(* IEC 61131-3 sources: daoli-st-library/DL_MathData (part 26) *)

(* ---- FC_DL_TimeDivChk.st ---- *)
(*
    FC_DL_TimeDivChk —— TIME 整数除法除零拦截与模长防御包装
    ------------------------------------------------------------------
    分类      : DL_MathData / TimeArith
    前缀      : FC_DL_
    版本      : 1.0.0
    溯源      : IEC 61131-3 标准语义的道莅防御性实现
                （内部委托平台内建函数，外围统一错误码/钳位/双语文档；
                  未复制任何闭源厂商源码，参考实现仅限 MIT/Apache 许可）
    平台      : 纯 IEC 61131-3，CODESYS / TwinCAT / InoProShop 通用
    作者      : 道莅代码库 · PLC编程专家（R16）
    ------------------------------------------------------------------
    功能说明  : TIME 整数除法：返回 tIn ÷ nDiv，TIME 算术委托 `÷` 运算符，
                不重实现任何时间运算内核；
                nDiv = 0 判为故障级 16#0001_02C7，返回 T#0S 且 bValid=FALSE（除零故障）；
                nDiv < 0 时取模长参与运算并置信息级 16#0001_01E6
                （TIME 无负语义，方向取模长，bError=FALSE、bValid=TRUE）；
                模长取负回绕防御：先将 INT 除子升位复制到 DINT 再取负，
                规避 INT 最小值 -32768 直接取负的回绕未定义行为；
                除法前已强制判定除子非零（nDiv = 0 分支提前拦截），满足除法前判除子红线；
                钳位方向：无钳位（除零故障拦截 / 负除子模长化记录）。
    错误码    : 16#0001_02C7 除数为 0（除零故障）——故障级，返回 T#0S
                16#0001_01E6 负除子输入，已按模长参与运算——信息级，正常防御
                16#0001_01E7 预留禁用（信息级，不得挪用）
                16#0001_02C8 预留禁用（故障级，不得挪用）
                16#0001_02C9 预留禁用（故障级，不得挪用）
    状态机    : R6 标注 N/A —— 本组件为纯函数无顺序状态机，无 CASE 可写，非法状态不可能出现，故以本节说明替代 ELSE 兜底
    修订记录  : 2026-11-16 v1.0.0 首次入库（R16）
*)
FUNCTION FC_DL_TimeDivChk : TIME
VAR_INPUT
    tIn  : TIME; // 输入时长（被除数） [ms] / input duration (dividend)
    nDiv : INT;  // 除子 [倍]，非 0，除零为故障 / divisor [x], nonzero, div-by-zero is a fault
END_VAR
VAR_OUTPUT
    eErr   : UDINT; // 错误码，0=正常 / error id, 0=ok
    bError : BOOL;  // 是否出错，eErr 非 0 时为 TRUE / error flag, TRUE when eErr is nonzero
    bValid : BOOL;  // 输出是否有效可用 / output valid flag
END_VAR
VAR CONSTANT
    DL_TIME_ZERO : TIME := T#0S; // TIME 零值（故障缺省返回） [ms] / TIME zero value (fault default return)
END_VAR
VAR
    nWiden : DINT; // 升位到 DINT 的除子副本 [倍] / divisor copy widened to DINT
    nAbs   : DINT; // 除子模长 [倍] / divisor magnitude
END_VAR

// 段 1｜返回值与错误状态预置 / segment 1, preset return value and error status
FC_DL_TimeDivChk := DL_TIME_ZERO; // 故障缺省返回 T#0S [ms] / fault default returns T#0S
eErr   := 0;     // 预置无错误 / preset no error
bError := FALSE; // 预置无故障 / preset no fault
bValid := FALSE; // 预置无效，通过除零闸后置位 / preset invalid, set TRUE after divide-by-zero guard

// 段 2｜除零故障闸 / segment 2, divide-by-zero fault guard
IF nDiv = 0 THEN
    FC_DL_TimeDivChk := DL_TIME_ZERO; // 故障级返回 T#0S [ms] / fault level returns T#0S
    eErr   := 16#0001_02C7;           // 除零故障码 / divide-by-zero fault id
    bError := TRUE;                   // 置故障标志 / set fault flag
    bValid := FALSE;                  // 输出无效 / output invalid
    RETURN;                           // 立即返回 / immediate return
END_IF

// 段 3｜除子模长整备（含取负回绕防御） / segment 3, divisor magnitude preparation with negation-wrap defense
nWiden := nDiv; // 先升位复制到 DINT / widen copy to DINT first
IF nDiv < 0 THEN
    nAbs := -nWiden; // DINT 域内取模长（规避 INT 最小值 -32768 取负回绕） / magnitude in DINT domain (avoids INT minimum -32768 negation wrap)
    eErr := 16#0001_01E6; // 信息级：负除子按模长处理（TIME 无负语义，方向取模长） / info level: negative divisor handled by magnitude (TIME has no negative semantics)
ELSE
    nAbs := nWiden; // 正除子模长即原值 / positive divisor, magnitude equals original
END_IF

// 段 4｜主体除法计算（末段） / segment 4, main division calculation (final)
FC_DL_TimeDivChk := tIn / nAbs; // 除子已判非零，模长参与委托 `÷` 运算符除法 / divisor checked nonzero, division via `÷` operator with magnitude
bError := FALSE; // 信息级模长化不置故障，除零分支已提前返回 / info-level magnitude never raises fault, divide-by-zero branch has returned
bValid := TRUE;  // 域内或模长化输出均有效可用 / in-domain or magnitude output is valid
END_FUNCTION

(* ---- FC_DL_TimeMulSat.st ---- *)
(*
    FC_DL_TimeMulSat —— TIME 整数乘法（乘数域闸 + 溢出饱和）
    ------------------------------------------------------------------
    分类      : DL_MathData / TimeArith
    前缀      : FC_DL_
    版本      : 1.0.0
    溯源      : IEC 61131-3 标准语义的道莅防御性实现
                （对照 IEC 61131-3 第 3 版 MUL_TIME 标准语义，委托平台内建 `*`
                  与 `/` 运算符，外围全部闸门 / 饱和 / 码位 / 双语文档 100% 自有；
                  clean-room 编写，未复制任何闭源厂商源码，参考实现仅限 MIT/Apache）
    平台      : 纯 IEC 61131-3，CODESYS 3.5 / TwinCAT 3 / InoProShop / Machine Expert 通用
    作者      : 道莅代码库 · PLC编程专家（R69 构建轮 · 批 1 · N1）
    ------------------------------------------------------------------
    功能说明  : TIME × 乘数。与库内既有 FC_DL_TimeScaleSat 的分工：ScaleSat 是
                「负乘子钳零、双乘子全放行」的宽松包装；本件是 MUL_TIME 的**严格域闸**
                版本——负乘子属于语义非法（时长无负语义）必须**禁入**并报故障级，
                乘数超 INT 正域上界（32767）同样禁入（防以超域乘子绕过溢出预判），
                只有域内合法乘子才进入乘法内核。
                溢出预判采用除法比较口径（R54 / 实战规则 6）：`tIn > MAX / nScale`，
                比较表达式中不出现乘 / 加运算符，命中即饱和夹 LTIME 上界并报信息级。
                乘数域上界反算依据（实战规则 9）：TIME 为 32 位毫秒容器
                （上限 4294967295 ms ≈ T#49D17H2M47S295MS），乘子上界取 32767（INT 正域）
                是为让 `MAX / nScale` 恒有整数解且不产生 0 除；乘子更大时预判式
                本身会因整数除法结果为 0 而把一切非零时长误判为溢出，故必须在域闸
                先行禁入，不得放大上界。
    错误码    : 16#0001_03F7 负乘子禁入（语义非法），输出 T#0S —— 故障级
                16#0001_03F8 乘子超上界 32767，输出 T#0S —— 故障级
                16#0001_04F6 乘法溢出，输出已饱和至 TIME 上界 —— 信息级，值可用
    码位总账  : 16#0001_03F7 / 03F8 用 ｜ 16#0001_04F6 用
    状态机    : R6 标注 N/A —— 纯函数无顺序状态机，无 CASE 可写，非法状态不可能出现
    采样约定  : 无定时器 / 无沿检测 / 无跨周期状态，结论与任务周期无关
    修订记录  : 2026-11-22 v1.0.0 首次入库（R69 构建轮 · 批 1 · N1）
*)
FUNCTION FC_DL_TimeMulSat : TIME
VAR_INPUT
    tIn     : TIME;                            // 被乘时长 [ms] / multiplicand duration [ms]
    diScale : DINT;                            // 乘数 [倍]，域 0..32767，负值与超上界禁入 / scale factor [x], domain 0..32767
END_VAR
VAR_OUTPUT
    eErr        : UDINT;                       // 错误码，0 = 正常 / error id, 0 = ok
    bError      : BOOL;                        // 故障标志，故障级码时为 TRUE / error flag, TRUE on fault level
    bValid      : BOOL;                        // 返回值可用（故障级为 FALSE）/ return usable, FALSE on fault level
    bSaturated  : BOOL;                        // 已饱和至 TIME 上界 / saturated at the TIME ceiling
END_VAR
VAR CONSTANT
    DL_TM_MAX   : TIME := T#49D17H2M47S295MS;  // 32 位 TIME 容器上限，等价 4294967295 ms [ms] / 32-bit TIME ceiling [ms]
    DL_TM_ZERO  : TIME := T#0S;                // TIME 零值（故障缺省返回） [ms] / TIME zero, the fault default
    DL_TM_SCALE_MAX : DINT := 32767;           // 乘数上界 [倍]，INT 正域上界（反算依据见头注释）/ scale ceiling [x]
    DL_TM_SCALE_MIN : DINT := 0;               // 乘数下界 [倍]，负值禁入 / scale floor [x]
END_VAR
VAR
    nScaleInt : INT;                           // 域内乘数（已过闸，可直接参与 TIME 运算）[倍] / in-domain scale as INT
END_VAR

// 段 1｜返回值与错误状态预置（实战规则 1① 四段式第一段）/ segment 1, preset return and status
FC_DL_TimeMulSat := DL_TM_ZERO;   // 故障缺省返回 T#0S [ms] / fault default returns T#0S
eErr       := 0;                  // 预置无错误 / preset no error
bError     := FALSE;              // 预置无故障 / preset no fault
bValid     := FALSE;              // 预置不可用，过闸后置位 / preset unusable, set TRUE after the gates
bSaturated := FALSE;              // 预置未饱和 / preset not saturated

// 段 2｜乘数域闸：负值禁入（语义非法）/ segment 2, scale domain gate, negative is refused
IF diScale < DL_TM_SCALE_MIN THEN
    eErr   := 16#0001_03F7;       // 故障级：负乘子禁入 / fault level: negative factor refused
    bError := TRUE;               // R45 配对置故障标志 / raise the error flag, paired with the code
    bValid := FALSE;              // 返回值不可用 / return unusable
    RETURN;                       // 出口，不触碰乘法内核 / exit, the kernel is never touched
END_IF

// 段 3｜乘数域闸：超上界禁入（防以超域乘子绕过溢出预判）/ segment 3, upper domain gate
IF diScale > DL_TM_SCALE_MAX THEN
    eErr   := 16#0001_03F8;       // 故障级：乘子超上界 / fault level: factor above the ceiling
    bError := TRUE;               // R45 配对 / paired with the code
    bValid := FALSE;              // 返回值不可用 / return unusable
    RETURN;                       // 出口 / exit
END_IF
nScaleInt := DINT_TO_INT(diScale);   // 域内乘数降为 INT（域已证 <= 32767，无窄化风险）[倍] / in-domain scale to INT

// 段 4｜零乘子：合法零乘，输出 T#0S 且无码（零乘不是错误）/ segment 4, legal zero multiply
IF nScaleInt = 0 THEN
    FC_DL_TimeMulSat := DL_TM_ZERO;   // 零乘结果 [ms] / zero product
    bValid := TRUE;                   // 零是可用结果 / zero is a usable result
    RETURN;                           // 出口 / exit
END_IF

// 段 5｜溢出预判（除法比较口径）+ 域内委托乘法内核 / segment 5, divide-compare pre-check then delegate
IF tIn > (DL_TM_MAX / nScaleInt) THEN
    FC_DL_TimeMulSat := DL_TM_MAX;    // 预判命中：饱和夹上界（除子 nScaleInt > 0 恒非零）[ms] / saturate to the ceiling
    eErr       := 16#0001_04F6;       // 信息级：乘法溢出已饱和 / info level: overflow saturated
    bSaturated := TRUE;               // 饱和标志供上层计量 / saturation flag for the caller
ELSE
    FC_DL_TimeMulSat := tIn * nScaleInt;   // 域内委托 `*` 运算符内核 [ms] / in-domain multiplication kernel
END_IF
bError := FALSE;   // 信息级饱和不置故障（饱和是防御而非故障）/ info-level saturation is a defence, not a fault
bValid := TRUE;    // 域内或饱和输出均可用 / usable in the in-domain and the saturated path
END_FUNCTION

(* ---- FC_DL_TimeRatioCalc.st ---- *)
(*
    FC_DL_TimeRatioCalc —— 两个 TIME 的无量纲比值
    ------------------------------------------------------------------
    分类      : DL_MathData / Convert
    前缀      : FC_DL_
    版本      : 1.0.0
    溯源      : 公开算术定义的道莅防御性实现（比值 = 分子时长 / 分母时长）；
                库内 FC_DL_TimeDivChk 只出整数毫秒商（小数全丢），本件用 LREAL 承载
                以保留 15 位有效数字；饱和限、取模长口径、错误分级、双语文档 100% 自有；
                clean-room 重写，未复制任何闭源厂商源码，参考实现仅限 MIT/Apache 许可
    平台      : 纯 IEC 61131-3，CODESYS V3.5+ / TwinCAT 3 / InoProShop 通用
    作者      : 道莅代码库 · PLC编程专家（R19）
    ------------------------------------------------------------------
    功能说明  : 计算节拍分析 / 稼动率 / 循环时间偏差 / 加速比所需的比值，可选 ×100 出百分比。
                核心防御：① 分母毫秒值为 0 是除零唯一出口（故障级 0321 早退，绝不进入除法）；
                ② 分母模长 < 1 ms 视为无意义分母，比值直接饱和到 fRatioSpan（1 ms 以下
                   的分母在任何现场都无意义，且会让比值爆炸）；
                ③ 输入为负时按模长参与运算（TIME 的平台符号语义不一致，方向差异
                   由本件统一吃掉），并置信息码 0402；
                ④ 比值超 fRatioSpan 双侧钳位，禁 NaN / ±INF 穿透；
                ⑤ 同一拍同时命中两条信息级时以 0403（饱和）为准，码位单值不可并列。
                职责边界：本件只出比值，不做时间加减、不做时基换算。
    错误码    : 16#0001_0402 分母模长 < 1 ms 或输入为负，已按模长运算/饱和——信息级，正常防御
                16#0001_0403 比值超 fRatioSpan 已钳位（bSaturated = TRUE）——信息级，正常防御
                16#0001_0321 分母为 0（除零）——故障级，返回 0.0 且 bValid = FALSE
                16#0001_0322 结果非有限（NaN / ±INF）或比值上限参数非法——故障级，返回 0.0
                16#0001_0323 预留禁用（故障级，不得挪用）
    码位总账  : 16#0001_0402 用 / 16#0001_0403 用 ｜ 16#0001_0321 用 / 16#0001_0322 用 / 16#0001_0323 预留
    状态机    : R6 标注 N/A —— 本组件为纯函数无顺序状态机，无 CASE 可写，非法状态不可能出现
    采样约定  : 本件无定时器、无沿检测；TIME 实参由调用方按自身时基给出，结论与任务周期无关。
    修订记录  : 2026-11-16 v1.0.0 首次入库（R19）
*)
FUNCTION FC_DL_TimeRatioCalc : LREAL
VAR_INPUT
    tNumerator      : TIME := T#0S;           // 分子时长 [ms]，域 -24 h~+24 h / numerator duration [ms], domain -24 h~+24 h
    tDenominator    : TIME := T#1S;           // 分母时长 [ms]，域 -24 h~+24 h，模长须 ≥ 1 ms / denominator duration [ms], domain -24 h~+24 h, magnitude >= 1 ms
    bAsPercent      : BOOL := FALSE;          // TRUE = 结果 ×100 输出百分比 [%] / TRUE multiplies the result by 100 to percent [%]
    fRatioSpan      : LREAL := 1.0E6;         // 比值饱和上限（作用在返回量上）[无量纲]，域 1.0~1.0E12 / ratio saturation span applied to the returned value [dimensionless], 1.0~1.0E12
END_VAR
VAR_OUTPUT
    eErr            : UDINT;                  // 错误码，0=正常 / error id, 0=ok
    bError          : BOOL;                   // 故障标志，eErr 为故障级时 TRUE / error flag, TRUE on fault-level eErr
    bValid          : BOOL;                   // 返回值是否可用 / return value valid flag
    fRatioAbs       : LREAL;                  // 比值绝对值（HMI 只看量级用）[无量纲] / absolute ratio for HMI magnitude view [dimensionless]
    bSaturated      : BOOL;                   // 比值已饱和到 fRatioSpan / ratio saturated to fRatioSpan
END_VAR
VAR CONSTANT
    DL_FLOAT_EPS        : REAL := 1.0E-6;     // 浮点判等容差 [无量纲] / float equality tolerance [dimensionless]
    DL_TR_MIN_DEN_MS    : LREAL := 1.0;       // 分母模长下限 [ms] / denominator magnitude lower bound [ms]
    DL_TR_PERCENT       : LREAL := 100.0;     // 百分比放大因子 [无量纲] / percent scale factor [dimensionless]
    DL_TR_SPAN_MIN      : LREAL := 1.0;       // 比值上限最小值 [无量纲] / minimum ratio span [dimensionless]
    DL_TR_SPAN_MAX      : LREAL := 1.0E12;    // 比值上限最大值 [无量纲] / maximum ratio span [dimensionless]
    DL_TR_INF_GUARD     : LREAL := 1.0E300;   // 非有限幅值判定阈值 [无量纲] / non-finite magnitude guard [dimensionless]
    DL_TR_ZERO          : LREAL := 0.0;       // 零值常量，避免裸字面量 [无量纲] / zero constant, avoids a bare literal [dimensionless]
END_VAR
VAR
    fNumAbs         : LREAL;                  // 分子模长 [ms] / numerator magnitude [ms]
    fDenAbs         : LREAL;                  // 分母模长 [ms] / denominator magnitude [ms]
    fSpanEff        : LREAL;                  // 生效比值上限，钳位后使用 [无量纲] / effective ratio span after clamping [dimensionless]
    fRatio          : LREAL;                  // 计算中的比值中间量 [无量纲] / ratio intermediate value [dimensionless]
    nDenMs          : DINT;                   // 分母毫秒整数形态，除零判定用 [ms] / denominator in integer milliseconds, used for the divide-by-zero gate [ms]
    bNegativeIn     : BOOL;                   // 输入存在负值时基的标志 / flag for negative time base inputs
END_VAR

// 段 1｜返回值与错误状态预置 / segment 1, preset return value and error status
FC_DL_TimeRatioCalc := DL_TR_ZERO;            // 故障缺省返回 0.0 / fault default returns zero
eErr := 0;                                    // 预置无错误 / preset no error
bError := FALSE;                              // 预置无故障 / preset no fault
bValid := FALSE;                              // 预置不可用，通过闸门后置位 / preset invalid, set TRUE after the gates
fRatioAbs := DL_TR_ZERO;                      // 量级输出先清零 / clear the magnitude output
bSaturated := FALSE;                          // 预置未饱和 / preset not saturated

// 段 2｜比值上限参数闸（非法上限等于比值域不存在，落入结果不可表示）/ segment 2, ratio span gate
fSpanEff := fRatioSpan;                       // 取入参副本，不改调用方数据 / copy the input, never modify caller data
IF (fSpanEff <> fSpanEff) OR (fSpanEff > DL_TR_INF_GUARD) OR (fSpanEff < -DL_TR_INF_GUARD) THEN
    eErr := 16#0001_0322;                     // 上限非有限即结果不可表示 / a non-finite span makes the result unrepresentable
    bError := TRUE;                           // 置故障标志 / raise the error flag
    RETURN;                                   // 故障级提前返回 / early return on fault
END_IF
IF fSpanEff < DL_TR_SPAN_MIN THEN
    fSpanEff := DL_TR_SPAN_MIN;               // 上限过小钳到 1.0，避免比值域退化 / clamp a too small span to 1.0
    eErr := 16#0001_0403;                     // 信息级：上限已钳位 / info level, the span has been clamped
ELSIF fSpanEff > DL_TR_SPAN_MAX THEN
    fSpanEff := DL_TR_SPAN_MAX;               // 上限过大钳到 1.0E12 / clamp an oversized span to 1.0E12
    eErr := 16#0001_0403;                     // 信息级：上限已钳位 / info level, the span has been clamped
END_IF

// 段 3｜除零唯一出口（先取整数毫秒判定，再进入浮点除法）/ segment 3, the only divide-by-zero exit
nDenMs := TIME_TO_DINT(tDenominator);         // 显式取分母毫秒整数，禁隐式换算 / take denominator milliseconds explicitly, no implicit cast
IF nDenMs = 0 THEN
    eErr := 16#0001_0321;                     // 除零故障码 / divide-by-zero fault id
    bError := TRUE;                           // 置故障标志 / raise the error flag
    bValid := FALSE;                          // 结果不可用 / result not usable
    RETURN;                                   // 故障级提前返回，绝不进入除法 / early return, the division is never executed
END_IF

// 段 4｜按模长参与运算（TIME 符号语义跨平台不一致，方向差异在此统一吃掉）/ segment 4, magnitudes only
fNumAbs := ABS(TIME_TO_LREAL(tNumerator));    // 分子模长 [ms] / numerator magnitude [ms]
fDenAbs := ABS(TIME_TO_LREAL(tDenominator));  // 分母模长 [ms] / denominator magnitude [ms]
bNegativeIn := (TIME_TO_DINT(tNumerator) < 0) OR (nDenMs < 0); // 负时基判定 / negative time base detection
IF bNegativeIn THEN
    eErr := 16#0001_0402;                     // 信息级：输入为负已按模长运算 / info level, negative inputs are handled by magnitude
END_IF

// 段 5｜分母过小闸：不足 1 ms 直接饱和，不做除法 / segment 5, tiny-denominator gate
IF fDenAbs < DL_TR_MIN_DEN_MS THEN
    fRatio := fSpanEff;                       // 过小分母直接给饱和值，规避比值爆炸 / jump straight to the span, avoid an exploding ratio
    bSaturated := TRUE;                       // 标记饱和 / flag the saturation
    eErr := 16#0001_0402;                     // 信息级：分母过小已饱和 / info level, tiny denominator saturated
ELSE
    fRatio := fNumAbs / fDenAbs;              // 分母模长 ≥ 1 ms，除法安全 / the denominator is at least 1 ms, the division is safe
    IF bAsPercent THEN
        fRatio := fRatio * DL_TR_PERCENT;     // 可选百分比放大 [%] / optional percent scaling [%]
    END_IF
END_IF

// 段 6｜结果非有限复检（NaN 穿透拦截）/ segment 6, non-finite recheck
IF (fRatio <> fRatio) OR (fRatio > DL_TR_INF_GUARD) OR (fRatio < -DL_TR_INF_GUARD) THEN
    eErr := 16#0001_0322;                     // 结果非有限故障码 / non-finite result fault id
    bError := TRUE;                           // 置故障标志 / raise the error flag
    bValid := FALSE;                          // 结果不可用 / result not usable
    FC_DL_TimeRatioCalc := DL_TR_ZERO;        // 明确返回 0.0 / return zero explicitly
    RETURN;                                   // 故障级提前返回 / early return on fault
END_IF

// 段 7｜饱和钳位（单侧上限，比值恒非负）/ segment 7, saturation clamp
IF fRatio > fSpanEff THEN
    fRatio := fSpanEff;                       // 钳到生效上限 / clamp to the effective span
    bSaturated := TRUE;                       // 标记饱和 / flag the saturation
    eErr := 16#0001_0403;                     // 信息级：超上限已钳位，与 0402 同拍时以本码为准 / info level, clamped; this id wins over 0402 in the same cycle
END_IF

// 段 8｜发布结果 / segment 8, publish the result
FC_DL_TimeRatioCalc := fRatio;                // 输出比值（含百分比放大） [无量纲] / publish the ratio incl. percent scaling [dimensionless]
fRatioAbs := fRatio;                          // 比值恒按模长运算，量级即本身 / the ratio is magnitude based, so the magnitude equals the value
bValid := TRUE;                               // 通过全部闸门，结果可用 / all gates passed, the result is usable
bError := FALSE;                              // 信息级不置故障 / info level never raises a fault
END_FUNCTION

(* ---- FC_DL_TimeScaleSat.st ---- *)
(*
    FC_DL_TimeScaleSat —— TIME 整数乘法溢出饱和防御包装
    ------------------------------------------------------------------
    分类      : DL_MathData / TimeArith
    前缀      : FC_DL_
    版本      : 1.0.0
    溯源      : IEC 61131-3 标准语义的道莅防御性实现
                （内部委托平台内建函数，外围统一错误码/钳位/双语文档；
                  未复制任何闭源厂商源码，参考实现仅限 MIT/Apache 许可）
    平台      : 纯 IEC 61131-3，CODESYS / TwinCAT / InoProShop 通用
    作者      : 道莅代码库 · PLC编程专家（R16）
    ------------------------------------------------------------------
    功能说明  : TIME 整数乘法：返回 tIn × nScale，TIME 算术委托 `×` 运算符，
                不重实现任何时间运算内核；
                nScale < 0 时防御性输出 T#0S 并置信息级 16#0001_01E5
                （TIME 无负语义，负乘子按钳零处理，bError=FALSE、bValid=TRUE）；
                nScale = 0 时输出 T#0S，无错误码（零乘合法）；
                溢出预判采用除法比较口径（规避「先算后判」红线）：
                nScale > 0 且 tIn > DL_TIME_MAX / nScale 时判乘法将溢出，
                直接饱和输出 DL_TIME_MAX，置信息级 16#0001_01E4；
                预判除法除子 nScale > 0 恒非零，满足除法前判除子红线；
                钳位方向：负乘子钳零 / 正乘子溢出钳上界 DL_TIME_MAX（双侧饱和语义）。
    错误码    : 16#0001_01E4 乘法结果超 TIME 上限，已饱和至 DL_TIME_MAX——信息级，正常防御
                16#0001_01E5 负乘子输入，已钳位输出 T#0S——信息级，正常防御
                16#0001_02C4 预留禁用（故障级，不得挪用）
                16#0001_02C5 预留禁用（故障级，不得挪用）
                16#0001_02C6 预留禁用（故障级，不得挪用）
    状态机    : R6 标注 N/A —— 本组件为纯函数无顺序状态机，无 CASE 可写，非法状态不可能出现，故以本节说明替代 ELSE 兜底
    修订记录  : 2026-11-16 v1.0.0 首次入库（R16）
*)
FUNCTION FC_DL_TimeScaleSat : TIME
VAR_INPUT
    tIn    : TIME; // 输入时长 [ms] / input duration
    nScale : INT;  // 乘子 [倍]，0~32767，负值输出钳 T#0s / scale factor [x], 0~32767, negative clamps output to T#0s
END_VAR
VAR_OUTPUT
    eErr   : UDINT; // 错误码，0=正常 / error id, 0=ok
    bError : BOOL;  // 是否出错，eErr 非 0 时为 TRUE / error flag, TRUE when eErr is nonzero
    bValid : BOOL;  // 输出是否有效可用 / output valid flag
END_VAR
VAR CONSTANT
    DL_TIME_MAX  : TIME := T#49D17H2M47S295MS; // 32 位 TIME 容器上限，等价 4294967295 ms [ms] / 32-bit TIME container ceiling, equals 4294967295 ms
    DL_TIME_ZERO : TIME := T#0S;               // TIME 零值（钳位目标） [ms] / TIME zero value (clamp target)
END_VAR

// 段 1｜返回值与错误状态预置 / segment 1, preset return value and error status
FC_DL_TimeScaleSat := DL_TIME_ZERO; // 故障缺省返回 T#0S [ms] / fault default returns T#0S
eErr   := 0;     // 预置无错误 / preset no error
bError := FALSE; // 预置无故障（本组件无故障级路径） / preset no fault (no fault-level path in this component)
bValid := FALSE; // 预置无效，通过乘子判定后置位 / preset invalid, set TRUE after factor check

// 段 2｜乘子符号判定 / segment 2, scale factor sign check
IF nScale < 0 THEN
    FC_DL_TimeScaleSat := DL_TIME_ZERO; // 负乘子钳位输出 T#0S（TIME 无负语义） / negative factor clamps output to T#0S (TIME has no negative semantics)
    eErr := 16#0001_01E5;               // 信息级：负乘子已钳零 / info level: negative factor clamped to zero
    bError := FALSE;                    // 信息级钳零不置故障 / info-level clamp never raises fault
    bValid := TRUE;                     // 钳零输出有效可用 / clamped output is valid
    RETURN;                             // 立即返回 / immediate return
ELSIF nScale = 0 THEN
    FC_DL_TimeScaleSat := DL_TIME_ZERO; // 零乘子输出 T#0S（零乘合法，无错误码） / zero factor yields T#0S (legal zero multiply, no error id)
    bError := FALSE;                    // 无故障 / no fault
    bValid := TRUE;                     // 输出有效可用 / output is valid
    RETURN;                             // 立即返回 / immediate return
END_IF

// 段 3｜除法比较溢出预判与主体乘法（末段） / segment 3, divide-compare overflow pre-check and main multiplication (final)
IF tIn > DL_TIME_MAX / nScale THEN
    FC_DL_TimeScaleSat := DL_TIME_MAX; // 溢出预判命中，饱和至上限（除子 nScale > 0 恒非零） / overflow pre-check hit, saturate to ceiling (divisor nScale > 0 guaranteed nonzero)
    eErr := 16#0001_01E4;              // 信息级：乘法溢出已饱和 / info level: multiplication overflow, saturated
ELSE
    FC_DL_TimeScaleSat := tIn * nScale; // 预判通过，域内委托 `×` 运算符乘法 / pre-check passed, in-domain multiplication via `×` operator
    eErr := 0; // 域内无错误 / in-domain, no error
END_IF
bError := FALSE; // 信息级饱和不置故障 / info-level saturation never raises fault
bValid := TRUE;  // 域内或饱和输出均有效可用 / in-domain or saturated output is valid
END_FUNCTION

(* ---- FC_DL_TimeSubSat.st ---- *)
(*
    FC_DL_TimeSubSat —— TIME 减法负差钳零防御包装
    ------------------------------------------------------------------
    分类      : DL_MathData / TimeArith
    前缀      : FC_DL_
    版本      : 1.0.0
    溯源      : IEC 61131-3 标准语义的道莅防御性实现
                （内部委托平台内建函数，外围统一错误码/钳位/双语文档；
                  未复制任何闭源厂商源码，参考实现仅限 MIT/Apache 许可）
    平台      : 纯 IEC 61131-3，CODESYS / TwinCAT / InoProShop 通用
    作者      : 道莅代码库 · PLC编程专家（R16）
    ------------------------------------------------------------------
    功能说明  : TIME 减法：返回 tA - tB（tA 为被减数、tB 为减数），TIME 算术
                委托 `-` 运算符，不重实现任何时间运算内核；
                tB > tA 时差为负，而 TIME 为无符号语义、负差跨平台未定义，
                故防御性钳位输出 T#0S 并置信息级 16#0001_01E2
                （bError=FALSE、bValid=TRUE，属正常防御）；
                钳位方向：仅下界单侧钳零（负差归 T#0S，不产生回绕）；
                本组件无故障级路径（减法运算不存在除法/非有限态故障源），
                故障三码位预留禁用。
    错误码    : 16#0001_01E2 减数为大，负差已钳位至 T#0S——信息级，正常防御
                16#0001_01E3 预留禁用（信息级，不得挪用）
                16#0001_02C1 预留禁用（故障级，不得挪用）
                16#0001_02C2 预留禁用（故障级，不得挪用）
                16#0001_02C3 预留禁用（故障级，不得挪用）
    状态机    : R6 标注 N/A —— 本组件为纯函数无顺序状态机，无 CASE 可写，非法状态不可能出现，故以本节说明替代 ELSE 兜底
    修订记录  : 2026-11-16 v1.0.0 首次入库（R16）
*)
FUNCTION FC_DL_TimeSubSat : TIME
VAR_INPUT
    tA : TIME; // 被减数 [ms] / minuend
    tB : TIME; // 减数 [ms] / subtrahend
END_VAR
VAR_OUTPUT
    eErr   : UDINT; // 错误码，0=正常 / error id, 0=ok
    bError : BOOL;  // 是否出错，eErr 非 0 时为 TRUE / error flag, TRUE when eErr is nonzero
    bValid : BOOL;  // 输出是否有效可用 / output valid flag
END_VAR
VAR CONSTANT
    DL_TIME_ZERO : TIME := T#0S; // TIME 零值（负差钳位目标） [ms] / TIME zero value (clamp target for negative difference)
END_VAR

// 段 1｜返回值与错误状态预置 / segment 1, preset return value and error status
FC_DL_TimeSubSat := DL_TIME_ZERO; // 故障缺省返回 T#0S [ms] / fault default returns T#0S
eErr   := 0;     // 预置无错误 / preset no error
bError := FALSE; // 预置无故障（本组件无故障级路径） / preset no fault (no fault-level path in this component)
bValid := FALSE; // 预置无效，通过负差判定后置位 / preset invalid, set TRUE after negative-difference check

// 段 2｜负差钳零判定与主体减法（末段） / segment 2, negative-difference clamp-to-zero check and main subtraction (final)
IF tB > tA THEN
    FC_DL_TimeSubSat := DL_TIME_ZERO; // 负差钳位至 T#0S（TIME 无符号语义，负差跨平台未定义） / negative difference clamped to T#0S (TIME is unsigned, negative difference is platform-undefined)
    eErr := 16#0001_01E2;             // 信息级：负差已钳零 / info level: negative difference clamped to zero
ELSE
    FC_DL_TimeSubSat := tA - tB; // 域内委托 `-` 运算符减法 / in-domain subtraction via `-` operator
    eErr := 0; // 域内无错误 / in-domain, no error
END_IF
bError := FALSE; // 信息级钳零不置故障 / info-level clamp never raises fault
bValid := TRUE;  // 域内或钳零输出均有效可用 / in-domain or clamped output is valid
END_FUNCTION

(* ---- FC_DL_TimeToDintMs.st ---- *)
(*
    FC_DL_TimeToDintMs —— TIME 到 DINT 毫秒防御转换（超域饱和）
    ------------------------------------------------------------------
    分类      : DL_MathData / TimeConv
    前缀      : FC_DL_
    版本      : 1.0.0
    溯源      : IEC 61131-3 标准语义的道莅防御性实现
                （接口语义由 IEC 61131-3 定义，内部委托平台内建 TIME_TO_DINT，
                  外围统一错误码 / 钳位 / 双语文档；clean-room 重写，
                  未复制任何闭源厂商源码，参考实现仅限 MIT/Apache 许可）
    平台      : 纯 IEC 61131-3，CODESYS / TwinCAT / InoProShop 通用
    作者      : 道莅代码库 · PLC编程专家（R17）
    ------------------------------------------------------------------
    功能说明  : 将 TIME 值防御性转换为 DINT 毫秒数并作为返回值输出，域内委托平台内建 TIME_TO_DINT；
                溢出预判先行：先在 TIME 域与 2147483647 ms（T#24D20H31M23S647MS）比较，
                超限直接饱和输出 2147483647 并置信息级 16#0001_01F2，
                严禁把超限值送进 TIME_TO_DINT（部分平台此时返回负值，静默翻转语义）；
                转换结果为负（负 TIME 或平台回绕）时钳 0 并置信息级 16#0001_01F3；
                钳位方向：上界饱和至 2147483647 ms，下界钳 0 ms；
                纯值类型域无 NaN/±INF 态，故无故障级路径（三个故障槽预留）。
    错误码    : 16#0001_01F2 输入超 DINT 毫秒域（> 2147483647 ms），已饱和——信息级，正常防御
                16#0001_01F3 转换结果为负（负 TIME 或平台回绕），已钳 0——信息级，正常防御
                16#0001_02D9 预留禁用（故障级，不得挪用）
                16#0001_02DA 预留禁用（故障级，不得挪用）
                16#0001_02DB 预留禁用（故障级，不得挪用）
    状态机    : R6 标注 N/A —— 本组件为纯函数无顺序状态机，无 CASE 可写，非法状态不可能出现，故以本节说明替代 ELSE 兜底
    修订记录  : 2026-11-16 v1.0.0 首次入库（R17）
*)
FUNCTION FC_DL_TimeToDintMs : DINT
VAR_INPUT
    tIn : TIME; // 待转换时间值，有效域 0 ms ~ 4294967295 ms [ms] / time value to convert, domain 0 ms .. 4294967295 ms [ms]
END_VAR
VAR_OUTPUT
    eErr   : UDINT; // 错误码，0=正常 / error id, 0=ok
    bError : BOOL;  // 是否出错，eErr 非 0 时为 TRUE / error flag, TRUE when eErr is nonzero
    bValid : BOOL;  // 输出是否有效可用 / output valid flag
END_VAR
VAR CONSTANT
    DL_TIME_DINT_MAX : TIME := T#24D20H31M23S647MS; // DINT 正域可承载的最大毫秒数 2147483647 ms [ms] / max ms a DINT can carry, 2147483647 ms [ms]
    DL_DINT_MAX_MS   : DINT := 2147483647;          // 上界饱和输出值 [ms] / upper saturation output [ms]
    DL_MS_MIN        : DINT := 0;                   // 下界钳位值（TIME 无负语义） [ms] / lower clamp, TIME has no negative semantics [ms]
END_VAR
VAR
    nOut : DINT; // 域内转换中间结果 [ms] / in-domain conversion intermediate [ms]
END_VAR

// 段 1｜返回值与错误状态预置 / segment 1, preset return value and error status
FC_DL_TimeToDintMs := DL_MS_MIN; // 故障缺省返回 0 ms（TIME 无负语义） [ms] / fault default 0 ms, TIME has no negative semantics [ms]
eErr   := 0;     // 预置无错误 / preset no error
bError := FALSE; // 预置无故障（本件无故障级路径） / preset no fault, no fault-level path here
bValid := FALSE; // 预置输出无效，通过上界预判后置位 / preset invalid, set TRUE after the upper-bound pre-check

// 段 2｜上界预判与饱和（先判后算，禁先转换） / segment 2, upper bound pre-check and saturation (compare before convert)
IF tIn > DL_TIME_DINT_MAX THEN // 在 TIME 域先比较，绝不让超限值进入内建转换 [ms] / compare in the TIME domain first, never let an oversized value reach the built-in conversion [ms]
    FC_DL_TimeToDintMs := DL_DINT_MAX_MS; // 饱和输出 DINT 正域上限 2147483647 ms [ms] / saturate to the DINT positive bound 2147483647 ms [ms]
    eErr := 16#0001_01F2;                 // 信息级：超 DINT 毫秒域已饱和，正常防御 / info level: beyond the DINT ms domain, saturated
    bError := FALSE;                      // 信息级不置故障 / info level never raises fault
    bValid := TRUE;                       // 饱和值本身有效可用 / the saturated value itself is valid
    RETURN;                               // 饱和即出口，不调用内建转换 / saturation is the exit, built-in conversion not called
END_IF

// 段 3｜域内委托转换与负值钳零（末段） / segment 3, in-domain delegated conversion and negative clamp (final)
nOut := TIME_TO_DINT(tIn); // 域内委托平台内建 TIME_TO_DINT [ms] / in-domain delegate to built-in TIME_TO_DINT [ms]
IF nOut < DL_MS_MIN THEN
    nOut := DL_MS_MIN;    // 负结果钳 0（负 TIME 或平台回绕，TIME 无负语义） [ms] / clamp negative results to 0, TIME has no negative semantics [ms]
    eErr := 16#0001_01F3; // 信息级：结果为负已钳零，正常防御 / info level: result was negative and clamped to zero
ELSE
    eErr := 0;            // 域内无错误 / in-domain, no error
END_IF
FC_DL_TimeToDintMs := nOut; // 输出钳位后的毫秒结果 [ms] / output the clamped millisecond result [ms]
bError := FALSE;            // 信息级不置故障 / info level never raises fault
bValid := TRUE;             // 域内或钳位后输出均有效可用 / in-domain or clamped output is valid
END_FUNCTION

(* ---- FC_DL_TimeToHmsString.st ---- *)
(*
    组件名称 : FC_DL_TimeToHmsString
    所属子库 : DL_MathData
    当前版本 : 1.0.0
    兼 容 性 : CODESYS V3.5+ / TwinCAT 3 / 汇川 InoProShop；仅依赖 Standard.library
    功能描述 : TIME 时长 → 'HH:MM:SS.mmm' 定宽文本，负时长统一带负号，并把总小时数单独出口供报表使用。
              取舍 ①：不委托 DINT_TO_STRING 补零 —— 各平台对「正数是否带前导空格」「负数符号位置」
              的实现互不相同（R79 家族），靠它拼定宽字段必出「_1:05:03」这类带空格的串。
              本件用数字字符表 MID 取值 + CONCAT 拼装，位数与字符完全由代码控制。
              取舍 ②：负数先取绝对值再分解，但 DINT_MIN 单独走哨兵分支 —— −(−2147483648) 在 DINT 域回绕成自身，
              直接取负会把「最大负时长」变成「最大正时长」且符号丢失；本件对下界显式夹到 DINT_MAX 并保留负号。
              取舍 ③：分解全程只用非负操作数 —— 取绝对值之后再 MOD/DIV，三平台的负数取余歧义从源头消失。
              取舍 ④：小时字段不设上限截断，只发宽度提示 —— TIME 上限约 596 小时，HMI 常见 2 位小时字段装不下，
              但截断小时会让时长错得无声无息，宁可超宽 + 信息码让上位机改字段宽度。
    开源溯源 : T2-1 LGF Converter 子族（只借「时长转定宽文本」这一行为定义）。码位、补零策略、负数口径、；本件为道莅 clean-room 防御性实现（仅借 LGF 分类事实/参数域/行为定义，零代码行与符号名复制）。
              分解顺序 100% 自有，零代码行与注释复制。
    本文件内含 : FUNCTION FC_DL_TimeToHmsString（单 POU，无配套类型）
    依 赖 : 无 DL_ 内部依赖；Standard.library: LEN / MID / CONCAT
    红线自检 : R1 ✓ 零全局变量与外部变量 ｜ R2 ✓ 零物理 IO 地址
              R3 ✓ 纯 IEC 61131-3 ｜ R4 ✓ 下界哨兵 + 小时域闸 + 分解操作数恒非负 + 输出长度自证
              R5 ✓ 全变量中英双语同行注释 ｜ R6 N/A 纯函数无顺序状态机，无 CASE 可写
              R7 N/A 无定时器、无沿检测实例 ｜ R8 ✓ 毫秒基数、字段宽度、小时上限全常量化
    错误码   : 16#0001_044E [信息级] 负时长已带负号输出，bValid = TRUE
               16#0001_044F [信息级] 小时超 99，HMI 两位小时字段装不下，bValid = TRUE
               16#0001_0393 [故障级] 分解中间量非法（小时超 999，理论不可达），返回 '00:00:00.000'，bValid = FALSE
               16#0001_0394 [故障级] 预留禁用（不得挪用）
               16#0001_0395 [故障级] 预留禁用（不得挪用）
    码位总账 : 16#0001_044E 用 / 16#0001_044F 用 ｜ 16#0001_0393 用 / 16#0001_0394 预留 / 16#0001_0395 预留
    遗留假设 : ① 本件依赖「平台 TIME 为 32 位有符号毫秒计数」这一口径（TIME_TO_DINT 与 TIME 同宽）。
              CODESYS / TwinCAT 3 默认如此，InoProShop 未实测；若某平台 TIME 换成 64 位 LTime 语义，
              小时上限与 DINT_MIN 哨兵都需重估。交付门槛：三平台各编译并跑 T#-1ms、T#-2147483648ms、
              T#596H 三个边界 —— 未实测，编译门槛未闭合。
              ② MID 参数序按 IEC 标准 MID(串, 长度, 位置)，与库内既有用法同序。
    修订历史 :
        2026-11-16  v1.0.0  首版，R21 批次 3 入库
*)
FUNCTION FC_DL_TimeToHmsString : STRING
VAR_INPUT
    tIn             : TIME;   // 待格式化时长，全域（含负值）[ms] / duration to format, negative values included [ms]
END_VAR
VAR_OUTPUT
    eErr            : UDINT;  // 错误码，0=正常；16#0001_04XX 信息级 / 16#0001_03XX 故障级 / error id, 0=ok
    bError          : BOOL;   // 故障级标志，eErr 落 16#0001_03XX 时为 TRUE / fault flag, TRUE on fault-level eErr
    bValid          : BOOL;   // 返回值是否可用 / result usable flag
    bNegative       : BOOL;   // 输入是否为负时长，输出串因此带前导负号 / TRUE when the input duration is negative and the text carries a minus sign
    nTotalHours     : DINT;   // 总小时数（分解后），供报表直接取用 [h] / total hours after the decomposition [h]
END_VAR
VAR
    nMs             : DINT;   // 时长的毫秒值，取绝对值后恒非负 [ms] / duration in milliseconds, non-negative after the magnitude step [ms]
    nHours          : DINT;   // 小时数 0~999 [h] / hours, 0..999 [h]
    nMinutes        : DINT;   // 分钟数 0~59 [min] / minutes, 0..59 [min]
    nSeconds        : DINT;   // 秒数 0~59 [s] / seconds, 0..59 [s]
    nMilli          : DINT;   // 毫秒数 0~999 [ms] / milliseconds, 0..999 [ms]
    sRet            : STRING; // 结果装配缓冲 [字符] / result assembly buffer [char]
    nDigits         : INT;    // 当前字段位数，用于补零循环 [位] / digits of the current field used by the padding loops [digit]
    nPos            : INT;    // 补零循环游标 [位] / padding loop cursor [digit]
END_VAR
VAR CONSTANT
    DL_MS_PER_SEC       : DINT := 1000;                  // 每秒毫秒数 [ms] / milliseconds per second [ms]
    DL_MS_PER_MIN       : DINT := 60000;                 // 每分毫秒数 [ms] / milliseconds per minute [ms]
    DL_MS_PER_HOUR      : DINT := 3600000;               // 每小时毫秒数 [ms] / milliseconds per hour [ms]
    DL_HMS_FIELD_WARN_H : DINT := 99;                    // HMI 常见两位小时字段上限 [h] / typical two digit hour field limit [h]
    DL_HMS_HOUR_MAX     : DINT := 999;                   // 三位小时字段上限，TIME 上限 596h 结构性不越此值 [h] / three digit hour field limit [h]
    DL_HMS_MS_MAX       : DINT := 999;                   // 毫秒字段上限 [ms] / millisecond field limit [ms]
    DL_HMS_MIN_MAX      : DINT := 60;                    // 分钟/秒的进位基数 [min] / radix of the minute and second fields [min]
    DL_HMS_DIGIT_TEN    : DINT := 10;                    // 十进制位数基数 [无量纲] / decimal digit radix [dimensionless]
    DL_HMS_DIGIT_HUND   : DINT := 100;                   // 百位基数 [无量纲] / hundreds radix [dimensionless]
    DL_DIGIT_TABLE      : STRING := '0123456789';        // 数字字符表，MID 位置 = 值 + 1 [字符] / digit table, the MID position is the value plus one [char]
    DL_HMS_COLON        : STRING := ':';                 // 时分秒分隔符 [字符] / hour-minute-second separator [char]
    DL_HMS_DOT          : STRING := '.';                 // 秒与毫秒分隔符 [字符] / second-millisecond separator [char]
    DL_HMS_MINUS        : STRING := '-';                 // 负号 [字符] / minus sign [char]
    DL_HMS_ZERO_TEXT    : STRING := '00:00:00.000';      // 故障回退串，长度恒 12 [字符] / fault fallback text with a constant length of twelve [char]
    DL_HMS_ZERO_CH      : STRING := '0';                 // 单个零字符，小时字段补位用 [字符] / single zero character used to pad the hour field [char]
    DL_HMS_ONE          : INT := 1;                      // 单位哨兵，MID 位置 1 基 [无量纲] / unity sentinel, MID is one based [dimensionless]
    DL_HMS_LEN_MIN      : INT := 12;                     // 最短合法长度（两位小时、无负号）[字符] / shortest legal length with two digit hours and no sign [char]
    DL_HMS_LEN_MAX      : INT := 14;                     // 最长合法长度（负号 + 三位小时）[字符] / longest legal length with a sign and three digit hours [char]
    DL_DINT_MIN         : DINT := -2147483648;           // DINT 下界，取负会回绕，必须单独拦 [ms] / DINT lower bound whose negation wraps around [ms]
    DL_DINT_MAX         : DINT := 2147483647;            // DINT 上界，下界夹到此值 [ms] / DINT upper bound used to clamp the lower bound case [ms]
    DL_DINT_ZERO        : DINT := 0;                     // 零哨兵 [ms] / zero sentinel [ms]
    DL_ERR_NONE         : UDINT := 16#0000_0000;         // 无故障 / no error
END_VAR

// 段 1｜返回值与错误状态预置 / segment 1, preset the return value and the error state
FC_DL_TimeToHmsString := DL_HMS_ZERO_TEXT;   // 故障缺省返回定宽零串 / fault default returns the fixed width zero text
eErr         := DL_ERR_NONE;                 // 预置无错误 / preset no error
bError       := FALSE;                       // 预置无故障 / preset no fault
bValid       := FALSE;                       // 预置结果不可用 / preset unusable
bNegative    := FALSE;                       // 预置非负 / preset non-negative
nTotalHours  := 0;                           // 预置小时 0 / preset the hours to zero
sRet         := '';                          // 缓冲清空 / clear the buffer

// 段 2｜取值与符号处理：下界单独夹，其余直接取负 / segment 2, magnitude step with an explicit lower bound branch
nMs := TIME_TO_DINT(tIn);                    // 毫秒口径，依赖平台 TIME 为 32 位毫秒（见遗留假设）/ millisecond reading, see the assumption note
IF nMs < DL_DINT_ZERO THEN
    bNegative := TRUE;                       // 标记负时长 / mark the negative duration
    eErr      := 16#0001_044E;               // 负时长已带负号输出（信息级，不置 bError）/ negative duration, info level
    IF nMs = DL_DINT_MIN THEN
        nMs := DL_DINT_MAX;                  // 下界取负会回绕，夹到上界（差 1ms，方向与符号均保留）/ negating the lower bound wraps, clamp instead
    ELSE
        nMs := -nMs;                         // 常规取绝对值 / usual magnitude
    END_IF
END_IF

// 段 3｜分解：操作数全程非负，MOD 无符号歧义 / segment 3, decomposition with non-negative operands only
nHours   := nMs / DL_MS_PER_HOUR;                          // 小时 / hours
nMinutes := (nMs MOD DL_MS_PER_HOUR) / DL_MS_PER_MIN;      // 分钟 / minutes
nSeconds := (nMs MOD DL_MS_PER_MIN) / DL_MS_PER_SEC;       // 秒 / seconds
nMilli   := nMs MOD DL_MS_PER_SEC;                         // 毫秒 / milliseconds
nTotalHours := nHours;                                     // 出口小时数 / publish the hours
IF nHours > DL_HMS_HOUR_MAX THEN
    eErr   := 16#0001_0393;              // 分解中间量非法（故障级，理论不可达）/ illegal intermediate, fault level, unreachable in theory
    bError := TRUE;                      // 置故障标志 / raise the fault flag
    RETURN;                              // 返回定宽零串 / return the fixed width zero text
END_IF
IF (nHours > DL_HMS_FIELD_WARN_H) AND (eErr = DL_ERR_NONE) THEN
    eErr := 16#0001_044F;                // 小时超 99 字段宽度提示（信息级）/ hour field too wide, info level
END_IF

// 段 4｜小时字段：最多三位，前导零按需省略 / segment 4, hour field with at most three digits and no superfluous zeros
IF bNegative THEN
    sRet := CONCAT(sRet, DL_HMS_MINUS);  // 负号前置 / the sign comes first
END_IF
IF nHours >= DL_HMS_DIGIT_HUND THEN
    sRet := CONCAT(sRet, MID(DL_DIGIT_TABLE, DL_HMS_ONE, DINT_TO_INT(nHours / DL_HMS_DIGIT_HUND) + DL_HMS_ONE));   // 百位 / hundreds digit
END_IF
IF nHours >= DL_HMS_DIGIT_TEN THEN
    sRet := CONCAT(sRet, MID(DL_DIGIT_TABLE, DL_HMS_ONE, DINT_TO_INT((nHours / DL_HMS_DIGIT_TEN) MOD DL_HMS_DIGIT_TEN) + DL_HMS_ONE));   // 十位 / tens digit
ELSE
    sRet := CONCAT(sRet, DL_HMS_ZERO_CH);   // 不足两位补零，保证 HH 定宽 / pad to two digits so the hour field keeps the HH width
END_IF
sRet := CONCAT(sRet, MID(DL_DIGIT_TABLE, DL_HMS_ONE, DINT_TO_INT(nHours MOD DL_HMS_DIGIT_TEN) + DL_HMS_ONE));   // 个位，恒输出 / units digit, always emitted
sRet := CONCAT(sRet, DL_HMS_COLON);      // 小时分隔符 / hour separator

// 段 5｜分钟与秒：两位定宽，逐位查表 / segment 5, minute and second fields, two digits each
sRet := CONCAT(sRet, MID(DL_DIGIT_TABLE, DL_HMS_ONE, DINT_TO_INT(nMinutes / DL_HMS_DIGIT_TEN) + DL_HMS_ONE));   // 分的十位 / minute tens
sRet := CONCAT(sRet, MID(DL_DIGIT_TABLE, DL_HMS_ONE, DINT_TO_INT(nMinutes MOD DL_HMS_DIGIT_TEN) + DL_HMS_ONE)); // 分的个位 / minute units
sRet := CONCAT(sRet, DL_HMS_COLON);      // 分隔符 / separator
sRet := CONCAT(sRet, MID(DL_DIGIT_TABLE, DL_HMS_ONE, DINT_TO_INT(nSeconds / DL_HMS_DIGIT_TEN) + DL_HMS_ONE));   // 秒的十位 / second tens
sRet := CONCAT(sRet, MID(DL_DIGIT_TABLE, DL_HMS_ONE, DINT_TO_INT(nSeconds MOD DL_HMS_DIGIT_TEN) + DL_HMS_ONE)); // 秒的个位 / second units
sRet := CONCAT(sRet, DL_HMS_DOT);        // 小数点 / decimal dot

// 段 6｜毫秒：三位定宽 / segment 6, millisecond field, three digits
sRet := CONCAT(sRet, MID(DL_DIGIT_TABLE, DL_HMS_ONE, DINT_TO_INT(nMilli / DL_HMS_DIGIT_HUND) + DL_HMS_ONE));   // 百位 / hundreds
sRet := CONCAT(sRet, MID(DL_DIGIT_TABLE, DL_HMS_ONE, DINT_TO_INT((nMilli / DL_HMS_DIGIT_TEN) MOD DL_HMS_DIGIT_TEN) + DL_HMS_ONE));   // 十位 / tens
sRet := CONCAT(sRet, MID(DL_DIGIT_TABLE, DL_HMS_ONE, DINT_TO_INT(nMilli MOD DL_HMS_DIGIT_TEN) + DL_HMS_ONE));   // 个位 / units

// 段 7｜出口长度自证：小时 ≤ 99 且非负为 12；带负号或三位小时为 13；两者兼有为 14 / segment 7, length self proof
nDigits := LEN(sRet);                    // 实际长度 / the actual length
IF (nDigits < DL_HMS_LEN_MIN) OR (nDigits > DL_HMS_LEN_MAX) THEN
    FC_DL_TimeToHmsString := DL_HMS_ZERO_TEXT;   // 长度异常回退定宽零串 / fall back to the fixed width zero text
    eErr   := 16#0001_0393;              // 格式装配异常按分解故障处置 / an assembly fault is reported as an intermediate fault
    bError := TRUE;                      // 置故障标志 / raise the fault flag
    RETURN;                              // bValid 保持 FALSE / bValid stays FALSE
END_IF

// 段 8｜出口 / segment 8, exit
FC_DL_TimeToHmsString := sRet;           // 输出定宽时间文本 / publish the fixed width time text
bValid := TRUE;                          // 结果可用 / the result is usable
END_FUNCTION

(* ---- FC_DL_TimeToLrealSec.st ---- *)
(*
    FC_DL_TimeToLrealSec —— TIME 到 LREAL 秒防御转换
    ------------------------------------------------------------------
    分类      : DL_MathData / TimeConv
    前缀      : FC_DL_
    版本      : 1.0.0
    溯源      : IEC 61131-3 标准语义的道莅防御性实现
                （接口语义由 IEC 61131-3 定义，内部委托平台内建 TIME_TO_LREAL，
                  外围统一错误码 / 钳位 / 双语文档；clean-room 重写，
                  未复制任何闭源厂商源码，参考实现仅限 MIT/Apache 许可）
    平台      : 纯 IEC 61131-3，CODESYS / TwinCAT / InoProShop 通用
    作者      : 道莅代码库 · PLC编程专家（R17）
    ------------------------------------------------------------------
    功能说明  : 将 TIME 值转换为 LREAL 秒数并作为返回值输出（节拍/速度/加速度算法的标准入口）；
                先委托平台内建 TIME_TO_LREAL 取毫秒数值，再除以常量 1000.0 得秒；
                除子为编译期常量 1000.0 恒非零，结构性满足除法前判除子非零红线；
                无上溢风险：TIME 域上限 4294967295 ms 远小于 2^53，LREAL 精确可表；
                负 TIME 照转不钳零（本件为观测语义，钳零会掩盖上游非法减法）并置信息级 16#0001_01F6；
                钳位方向：无钳位（仅记录负值，输出值与输入严格等价）。
    错误码    : 16#0001_01F6 负 TIME 输入（照转不钳零，仅记录）——信息级，正常防御
                16#0001_01F7 预留禁用（信息级，不得挪用）
                16#0001_02DF 预留禁用（故障级，不得挪用）
                16#0001_02E0 预留禁用（故障级，不得挪用）
                16#0001_02E1 预留禁用（故障级，不得挪用）
    状态机    : R6 标注 N/A —— 本组件为纯函数无顺序状态机，无 CASE 可写，非法状态不可能出现，故以本节说明替代 ELSE 兜底
    修订记录  : 2026-11-16 v1.0.0 首次入库（R17）
*)
FUNCTION FC_DL_TimeToLrealSec : LREAL
VAR_INPUT
    tIn : TIME; // 待转换时间值，有效域 0 ms ~ 4294967295 ms [ms] / time value to convert, domain 0 ms .. 4294967295 ms [ms]
END_VAR
VAR_OUTPUT
    eErr   : UDINT; // 错误码，0=正常 / error id, 0=ok
    bError : BOOL;  // 是否出错，eErr 非 0 时为 TRUE / error flag, TRUE when eErr is nonzero
    bValid : BOOL;  // 输出是否有效可用 / output valid flag
END_VAR
VAR CONSTANT
    DL_MS_PER_SEC : LREAL := 1000.0; // 毫秒/秒换算除子（编译期常量，恒非零） [ms/s] / ms-per-second divisor, compile-time constant, never zero [ms/s]
    DL_LREAL_ZERO : LREAL := 0.0;    // 返回值预置零（本件无故障路径，仅作预置约定） [s] / preset zero, no fault path in this component [s]
END_VAR
VAR
    fMsL : LREAL; // 毫秒数值（LREAL 承载） [ms] / millisecond value carried in LREAL [ms]
END_VAR

// 段 1｜返回值与错误状态预置 / segment 1, preset return value and error status
FC_DL_TimeToLrealSec := DL_LREAL_ZERO; // 故障缺省预置 0.0 s（本件无故障级路径） [s] / preset 0.0 s, no fault-level path in this component [s]
eErr   := 0;     // 预置无错误 / preset no error
bError := FALSE; // 预置无故障（本件无故障级路径） / preset no fault, no fault-level path here
bValid := FALSE; // 预置输出无效，通过数值整备后置位 / preset invalid, set TRUE after value preparation

// 段 2｜毫秒数值整备与负值记录 / segment 2, millisecond preparation and negative value recording
fMsL := TIME_TO_LREAL(tIn); // 委托平台内建 TIME_TO_LREAL 取毫秒数值 [ms] / delegate to built-in TIME_TO_LREAL for the millisecond value [ms]
IF fMsL < 0.0 THEN
    eErr := 16#0001_01F6; // 信息级：负 TIME 照转不钳零，仅记录（钳零会掩盖上游非法减法） / info level: negative TIME passed through and recorded only, clamping would hide an illegal upstream subtraction
ELSE
    eErr := 0;            // 非负时间无错误 / non-negative time, no error
END_IF

// 段 3｜毫秒转秒（末段） / segment 3, milliseconds to seconds (final)
FC_DL_TimeToLrealSec := fMsL / DL_MS_PER_SEC; // 除子为编译期常量 1000.0，恒非零 [s] / divisor is the compile-time constant 1000.0, never zero [s]
bError := FALSE;                              // 信息级不置故障 / info level never raises fault
bValid := TRUE;                               // 域内输出有效可用（负值亦有效，仅附信息码） / output is valid in-domain, including recorded negatives
END_FUNCTION

(* ---- FC_DL_TodAddWrap.st ---- *)
(*
    FC_DL_TodAddWrap —— TOD 加 TIME 偏移的午夜回绕加法
    ------------------------------------------------------------------
    分类      : DL_MathData / TimeArith
    前缀      : FC_DL_
    版本      : 1.0.0
    溯源      : IEC 61131-3 标准语义的道莅防御性实现（TOD + TIME → TOD，跨零点回绕）；
                委托平台内建 TOD_TO_DINT / TIME_TO_DINT / DINT_TO_TOD 完成显式换算，
                本件不重实现时间算术内核；
                偏移模长闸、回绕归一、回绕圈数回告、错误分级与码位 100% 自有；
                clean-room 重写，未复制任何闭源厂商源码，参考实现仅限 MIT/Apache 许可
    平台      : 纯 IEC 61131-3，CODESYS V3.5+ / TwinCAT 3 / InoProShop 通用
    作者      : 道莅代码库 · PLC编程专家（R20）
    ------------------------------------------------------------------
    功能说明  : 排程偏移、班次推算、延时启动时刻这类场景要把当日时刻加/减一段时间，
                结果必须落在同一日的 TOD 域内（跨零点即回绕）。与 DINT 毫秒加法件的
                本质区别是：TOD 域是环形的，回绕不是溢出而是正常语义。
                核心防御：① 全程显式标准转换（TOD_TO_DINT / TIME_TO_DINT），禁隐式赋值，
                   时间位型在不同平台的隐式转换口径不一致；
                ② 回绕归一**禁用取模**：负数取余在三种平台上分别可能是截断、向下取整或
                   实现未定义（R11 RolloverCounter 纪律），本件改条件加减；
                ③ 单次条件加减即可覆盖全域，条件是结构性成立的：段 2 已把偏移模长收到
                   一日以内、段 3 已把基准时刻收到 [0, 一日)，故 nSum 必落在
                   (−一日, 2×一日) 的开区间内，一次加或减必然落域，无需循环；
                ④ 偏移模长 ≥ 一日直接升故障级 034E：排程偏移不存在跨日以上的语义，
                   宁报不用——回绕圈数虽可算，但调用方拿到的多半不是他要的东西；
                ⑤ 回绕发生即置 bWrapped 与带符号的 nWrapCircles，方向可查；
                ⑥ 归一后再断言一次落域（034F），防平台时间位型异常。
                职责边界：两 TOD 之差（跨零点为正）归 FC_DL_TodDiffWrap；
                DINT 毫秒 → TOD 的纯转换归 FC_DL_DintMsToTod；本件只管带偏移的回绕加法。
    编译门槛  : 主路径依赖平台内建 TOD_TO_DINT（TOD 毫秒口径）、TIME_TO_DINT（TIME 毫秒口径）、
                DINT_TO_TOD。三平台标准库均提供；若某平台 TOD 以 32 位毫秒承载而 TIME 以
                64 位承载，段 3 的落域断言会拦下 TIME_TO_DINT 的高位截断，不会静默出错。
    错误码    : 16#0001_0420 发生午夜回绕（bWrapped 与 nWrapCircles 可查）——信息级，值可用
                16#0001_0421 预留禁用（信息级，不得挪用）
                16#0001_034E 偏移模长超一日，超出本件收窄域——故障级，返回 TOD 零点
                16#0001_034F 合成路径中间量非域（基准时刻或归一后结果越界）——故障级，返回 TOD 零点
                16#0001_0350 预留禁用（故障级，不得挪用）
    码位总账  : 16#0001_0420 用 / 16#0001_0421 预留 ｜ 16#0001_034E 用 / 16#0001_034F 用 / 16#0001_0350 预留
    状态机    : R6 标注 N/A —— 本组件为纯函数无顺序状态机，无 CASE 可写，非法状态不可能出现
    采样约定  : 本件无定时器、无沿检测、无状态；单拍纯计算，结论与任务周期无关。
    修订记录  : 2026-11-16 v1.0.0 首次入库（R20）
*)
FUNCTION FC_DL_TodAddWrap : TOD
VAR_INPUT
    todIn            : TOD;                   // 当日基准时刻 [时刻]，有效域 00:00:00.000~23:59:59.999 / base time of day [time of day], valid domain 00:00:00.000 to 23:59:59.999
    tOffset          : TIME;                  // 时刻偏移，可正可负 [ms]，本件收窄到模长 < 一日 / offset, signed [ms], narrowed to less than one day
END_VAR
VAR_OUTPUT
    eErr             : UDINT;                 // 错误码，0=正常 / error id, 0=ok
    bError           : BOOL;                  // 故障标志，eErr 为故障级时 TRUE / error flag, TRUE on fault-level eErr
    bValid           : BOOL;                  // 返回值是否可用（故障级为 FALSE）/ return usable, FALSE on fault level
    bWrapped         : BOOL;                  // 本拍发生午夜回绕 / a midnight wrap happened in this cycle
    nWrapCircles     : INT;                   // 回绕圈数，正向 +1、负向 −1，未回绕为 0 [圈] / wrap circles, +1 forward, −1 backward, 0 when no wrap [circle]
END_VAR
VAR CONSTANT
    DL_TOD_DAY_MS    : DINT := 86400000;      // 当日毫秒数 [ms/日] / milliseconds per day [ms/day]
    DL_TOD_DAY_NEG_MS : DINT := -86400000;    // 当日毫秒数的负值，负向闸门用 [ms/日] / negative milliseconds per day used by the backward gate [ms/day]
    DL_DINT_ZERO     : DINT := 0;             // 有符号零常量，避免裸字面量 [ms] / signed zero constant [ms]
    DL_WRAP_POS      : INT := 1;              // 正向回绕圈数 [圈] / positive wrap circle [circle]
    DL_WRAP_NEG      : INT := -1;             // 负向回绕圈数 [圈] / negative wrap circle [circle]
    DL_WRAP_NONE     : INT := 0;              // 未回绕时的圈数 [圈] / the circle count when nothing wrapped [circle]
    DL_TOD_ZERO      : TOD := TOD#00:00:00;   // 故障缺省返回的当日零点 / the midnight instant returned on faults
END_VAR
VAR
    nBase            : DINT;                  // 基准时刻毫秒中间量 [ms] / base time of day in milliseconds [ms]
    nOff             : DINT;                  // 偏移毫秒中间量 [ms] / offset in milliseconds [ms]
    nSum             : DINT;                  // 求和与归一中间量 [ms] / sum and normalisation intermediate [ms]
END_VAR

// 段 1｜返回值与错误状态预置 / segment 1, preset return value and error status
FC_DL_TodAddWrap := DL_TOD_ZERO;              // 故障缺省返回当日零点 / fault default returns midnight
eErr := 0;                                    // 预置无错误 / preset no error
bError := FALSE;                              // 预置无故障 / preset no fault
bValid := FALSE;                              // 预置不可用，通过闸门后置位 / preset invalid, set TRUE after the gates
bWrapped := FALSE;                            // 预置未回绕 / preset no wrap
nWrapCircles := DL_WRAP_NONE;                 // 预置回绕圈数 0 [圈] / preset zero wrap circles [circle]
nSum := DL_DINT_ZERO;                         // 归一中间量清零 / clear the normalisation intermediate

// 段 2｜偏移模长闸：跨日以上的偏移不在本件语义内，先判后算 / segment 2, offset magnitude gate
nOff := TIME_TO_DINT(tOffset);                // TIME → 毫秒，显式标准转换 [ms] / explicit standard conversion from TIME to milliseconds [ms]
IF (nOff >= DL_TOD_DAY_MS) OR (nOff <= DL_TOD_DAY_NEG_MS) THEN
    eErr := 16#0001_034E;                     // 故障级：偏移模长超一日 / fault level, the offset magnitude reaches one day
    bError := TRUE;                           // 置故障标志 / raise the error flag
    bValid := FALSE;                          // 返回值不可用 / flag the return as unusable
    FC_DL_TodAddWrap := DL_TOD_ZERO;          // 确定缺省值：当日零点 / deterministic default of midnight
    RETURN;                                   // 出口，不触碰时间合成 / exit, no time synthesis happens
END_IF

// 段 3｜基准时刻域闸：TOD 必须落在 [0, 一日) / segment 3, base time domain gate
nBase := TOD_TO_DINT(todIn);                  // TOD → 毫秒，显式标准转换 [ms] / explicit standard conversion from TOD to milliseconds [ms]
IF (nBase < DL_DINT_ZERO) OR (nBase >= DL_TOD_DAY_MS) THEN
    eErr := 16#0001_034F;                     // 故障级：合成路径中间量非域 / fault level, an intermediate left its domain
    bError := TRUE;                           // 置故障标志 / raise the error flag
    bValid := FALSE;                          // 返回值不可用 / flag the return as unusable
    FC_DL_TodAddWrap := DL_TOD_ZERO;          // 确定缺省值：当日零点 / deterministic default of midnight
    RETURN;                                   // 出口 / exit
END_IF

// 段 4｜求和：两操作数均已收窄，DINT 加法结构性不溢出 / segment 4, summation, structurally overflow free
nSum := nBase + nOff;                         // 基准毫秒 + 偏移毫秒 [ms] / base milliseconds plus offset milliseconds [ms]

// 段 5｜回绕归一：条件加减，禁用取模（R11 纪律）/ segment 5, wrap normalisation by conditional add and subtract
IF nSum >= DL_TOD_DAY_MS THEN
    nSum := nSum - DL_TOD_DAY_MS;             // 正向回绕减一日 [ms] / forward wrap, subtract one day [ms]
    nWrapCircles := DL_WRAP_POS;              // 圈数 +1 [圈] / one forward circle [circle]
    bWrapped := TRUE;                         // 标记回绕 / flag the wrap
    eErr := 16#0001_0420;                     // 信息级：发生午夜回绕 / info level, a midnight wrap happened
ELSIF nSum < DL_DINT_ZERO THEN
    nSum := nSum + DL_TOD_DAY_MS;             // 负向回绕加一日 [ms] / backward wrap, add one day [ms]
    nWrapCircles := DL_WRAP_NEG;              // 圈数 −1 [圈] / one backward circle [circle]
    bWrapped := TRUE;                         // 标记回绕 / flag the wrap
    eErr := 16#0001_0420;                     // 信息级：发生午夜回绕 / info level, a midnight wrap happened
END_IF

// 段 6｜归一后落域断言（双保险，防平台时间位型异常）/ segment 6, post-normalisation domain assertion
IF (nSum < DL_DINT_ZERO) OR (nSum >= DL_TOD_DAY_MS) THEN
    eErr := 16#0001_034F;                     // 故障级：归一后仍越界，平台时间位型异常 / fault level, still out of domain after normalisation
    bError := TRUE;                           // 置故障标志 / raise the error flag
    bValid := FALSE;                          // 返回值不可用 / flag the return as unusable
    FC_DL_TodAddWrap := DL_TOD_ZERO;          // 确定缺省值：当日零点 / deterministic default of midnight
    RETURN;                                   // 出口 / exit
END_IF

// 段 7｜发布结果 / segment 7, publish the result
FC_DL_TodAddWrap := DINT_TO_TOD(nSum);        // 毫秒 → 当日时刻 [时刻] / milliseconds back to a time of day [time of day]
bValid := TRUE;                               // 域内与回绕均可用 / usable in domain and after a wrap
bError := FALSE;                              // 信息级不置故障 / info level never raises a fault
END_FUNCTION

(* ---- FC_DL_TodDiffWrap.st ---- *)
(*
    FC_DL_TodDiffWrap —— 两 TOD 之差（跨零点为正）
    ------------------------------------------------------------------
    分类      : DL_MathData / TimeArith
    前缀      : FC_DL_
    版本      : 1.0.0
    溯源      : IEC 61131-3 标准语义的道莅防御性实现（两个当日时刻的区间时长，跨零点折算）；
                委托平台内建 TOD_TO_DINT / DINT_TO_TIME 完成显式换算，本件不重实现时间算术内核；
                跨零点判定、单次折算、跨零点标志与码位 100% 自有；
                clean-room 重写，未复制任何闭源厂商源码，参考实现仅限 MIT/Apache 许可
    平台      : 纯 IEC 61131-3，CODESYS V3.5+ / TwinCAT 3 / InoProShop 通用
    作者      : 道莅代码库 · PLC编程专家（R20）
    ------------------------------------------------------------------
    功能说明  : 班次工时、节拍间隔、夜间保温时段时长的高频口径：给两个当日时刻，
                求「从前者走到后者」的时长；后者小于前者即视为跨零点，按加一日折算，
                结果恒为非负。与 FC_DL_TodAddWrap 的加偏移语义互补。
                核心防御：① 差值后判定为负才加一日，且**只加一次**——判据是结构性的：
                   TOD 类型值域为 [0, 一日)，两值之差的模长必小于一日，故单次折算必然落域，
                   不需要循环也不需要取模（负数取余的三平台口径不一致，R11 纪律）；
                ② 本件五槽中信息 1 槽使用、故障 3 槽按规格预留禁用——域外输入在此件的
                   类型域上不可表达（TOD 值域由类型系统保证），故不设故障出口，
                   也不为「不存在的越界」虚构码位；
                ③ 跨零点事件用 bCrossMidnight 回告，HMI 可据此区分「同日间隔」与
                   「跨零点间隔」，否则 2 小时的结果看不出是凌晨还是傍晚来的；
                ④ 全程显式标准转换，禁隐式赋值。
                职责边界：时刻加偏移归 FC_DL_TodAddWrap；窗内判定归 FB_DL_TimeWindowCheck
                （它不提供原子差值）；本件只管两时刻的区间时长。
    编译门槛  : 主路径依赖平台内建 TOD_TO_DINT（毫秒口径）与 DINT_TO_TIME。
                三平台标准库均提供；结果上限 86399999 ms 恒落在 TIME 正域内，
                不存在 TIME 位型截断风险。
    错误码    : 16#0001_0422 跨零点区间（已按加一日折算，bCrossMidnight 可查）——信息级，值可用
                16#0001_0423 预留禁用（信息级，不得挪用）
                16#0001_0351 预留（故障级，不得挪用）
                16#0001_0352 预留禁用（故障级，不得挪用）
                16#0001_0353 预留禁用（故障级，不得挪用）
    码位总账  : 16#0001_0422 用 / 16#0001_0423 预留 ｜ 16#0001_0351 预留 / 16#0001_0352 预留 / 16#0001_0353 预留
    状态机    : R6 标注 N/A —— 本组件为纯函数无顺序状态机，无 CASE 可写，非法状态不可能出现
    采样约定  : 本件无定时器、无沿检测、无状态；单拍纯计算，结论与任务周期无关。
    修订记录  : 2026-11-16 v1.0.0 首次入库（R20）
*)
FUNCTION FC_DL_TodDiffWrap : TIME
VAR_INPUT
    todEarlier       : TOD;                   // 区间起点时刻 [时刻]，有效域 00:00:00.000~23:59:59.999 / start of the interval [time of day]
    todLater         : TOD;                   // 区间终点时刻 [时刻]，小于起点即视为跨零点 / end of the interval [time of day], earlier than the start means a midnight crossing
END_VAR
VAR_OUTPUT
    eErr             : UDINT;                 // 错误码，0=正常 / error id, 0=ok
    bError           : BOOL;                  // 故障标志，本件无故障级出口，恒为 FALSE / error flag, always FALSE here as no fault exit exists
    bValid           : BOOL;                  // 返回值是否可用（本件恒为 TRUE）/ return usable, always TRUE here
    bCrossMidnight   : BOOL;                  // 区间跨零点判定 / the interval crosses midnight
END_VAR
VAR CONSTANT
    DL_TOD_DAY_MS    : DINT := 86400000;      // 当日毫秒数 [ms/日] / milliseconds per day [ms/day]
    DL_DINT_ZERO     : DINT := 0;             // 有符号零常量，避免裸字面量 [ms] / signed zero constant [ms]
    DL_TIME_ZERO     : TIME := T#0s;          // 零时长，缺省返回 / zero duration returned by default
END_VAR
VAR
    nFrom            : DINT;                  // 起点时刻毫秒 [ms] / start instant in milliseconds [ms]
    nTo              : DINT;                  // 终点时刻毫秒 [ms] / end instant in milliseconds [ms]
    nDiff            : DINT;                  // 区间时长中间量，可为负 [ms] / interval duration intermediate, possibly negative [ms]
END_VAR

// 段 1｜返回值与错误状态预置 / segment 1, preset return value and error status
FC_DL_TodDiffWrap := DL_TIME_ZERO;            // 缺省返回零时长 / default returns a zero duration
eErr := 0;                                    // 预置无错误 / preset no error
bError := FALSE;                              // 本件无故障级出口，恒 FALSE / no fault exit exists, always FALSE
bValid := FALSE;                              // 预置不可用，通过闸门后置位 / preset invalid, set TRUE after the gates
bCrossMidnight := FALSE;                      // 预置未跨零点 / preset no midnight crossing
nDiff := DL_DINT_ZERO;                        // 中间量清零 / clear the intermediate

// 段 2｜取值：两时刻各做一次显式标准转换 / segment 2, both instants are converted explicitly
nFrom := TOD_TO_DINT(todEarlier);             // 起点毫秒 [ms] / start instant in milliseconds [ms]
nTo := TOD_TO_DINT(todLater);                 // 终点毫秒 [ms] / end instant in milliseconds [ms]

// 段 3｜求差：模长必小于一日的结构性事实来自 TOD 类型值域 / segment 3, difference bounded by one day
nDiff := nTo - nFrom;                         // 有符号区间差 [ms] / signed interval difference [ms]

// 段 4｜跨零点单次折算（禁取模，只加一次）/ segment 4, single midnight conversion without any modulo
IF nDiff < DL_DINT_ZERO THEN
    nDiff := nDiff + DL_TOD_DAY_MS;           // 负差值加一日折算为正 [ms] / add one day so the value becomes positive [ms]
    bCrossMidnight := TRUE;                   // 标记跨零点 / flag the midnight crossing
    eErr := 16#0001_0422;                     // 信息级：跨零点区间已折算 / info level, the interval crossed midnight and was converted
END_IF

// 段 5｜发布结果 / segment 5, publish the result
FC_DL_TodDiffWrap := DINT_TO_TIME(nDiff);     // 毫秒 → 时长 [ms] / milliseconds back to a duration [ms]
bValid := TRUE;                               // 折算后恒落 TIME 正域 / always inside the positive TIME domain after the conversion
bError := FALSE;                              // 信息级不置故障（双保险）/ info level never raises a fault, second line of defence
END_FUNCTION

(* ---- FC_DL_TodToDintMs.st ---- *)
(*
    FC_DL_TodToDintMs —— TOD 到当日毫秒偏移防御转换
    ------------------------------------------------------------------
    分类      : DL_MathData / TimeConv
    前缀      : FC_DL_
    版本      : 1.0.0
    溯源      : IEC 61131-3 标准语义的道莅防御性实现
                （接口语义由 IEC 61131-3 定义，内部委托平台内建 TOD_TO_TIME 与 TIME_TO_DINT，
                  外围统一错误码 / 钳位 / 双语文档；clean-room 重写，
                  未复制任何闭源厂商源码，参考实现仅限 MIT/Apache 许可）
    平台      : 纯 IEC 61131-3，CODESYS / TwinCAT / InoProShop 通用
    作者      : 道莅代码库 · PLC编程专家（R17）
    ------------------------------------------------------------------
    功能说明  : 将 TOD（当日时刻）转换为当日 0 点起的毫秒偏移并作为返回值输出，
                内部委托标准转换链 TOD_TO_TIME 再 TIME_TO_DINT，不自行按小时/分/秒累加
                （自实现累加会把时区、闰秒、平台 TOD 精度差异一并写进业务代码）；
                结果越出 0 ~ 86399999 ms 时按方向钳位并置信息级 16#0001_01FA；
                钳位方向：下界 0 ms，上界 86399999 ms（24h − 1 ms）；
                纯值类型域无 NaN/±INF 态，故无故障级路径（三个故障槽预留）；
                交付门槛：本件因依赖 TOD_TO_TIME 链，须在 CODESYS / TwinCAT / InoProShop 三平台各编译验证一次。
    错误码    : 16#0001_01FA TOD 转换结果越出 0 ~ 86399999 ms，已按方向钳位——信息级，正常防御
                16#0001_01FB 预留禁用（信息级，不得挪用）
                16#0001_02E5 预留禁用（故障级，不得挪用）
                16#0001_02E6 预留禁用（故障级，不得挪用）
                16#0001_02E7 预留禁用（故障级，不得挪用）
    状态机    : R6 标注 N/A —— 本组件为纯函数无顺序状态机，无 CASE 可写，非法状态不可能出现，故以本节说明替代 ELSE 兜底
    修订记录  : 2026-11-16 v1.0.0 首次入库（R17）
*)
FUNCTION FC_DL_TodToDintMs : DINT
VAR_INPUT
    todIn : TOD; // 当日时刻，有效域 00:00:00 ~ 23:59:59.999 [ms since 00:00:00] / time of day, domain 00:00:00 .. 23:59:59.999 [ms since midnight]
END_VAR
VAR_OUTPUT
    eErr   : UDINT; // 错误码，0=正常 / error id, 0=ok
    bError : BOOL;  // 是否出错，eErr 非 0 时为 TRUE / error flag, TRUE when eErr is nonzero
    bValid : BOOL;  // 输出是否有效可用 / output valid flag
END_VAR
VAR CONSTANT
    DL_TOD_MAX_MS : DINT := 86399999; // 当日毫秒上界（24h − 1 ms） [ms] / day upper bound, 24h minus 1 ms [ms]
    DL_TOD_MIN_MS : DINT := 0;        // 当日毫秒下界 [ms] / day lower bound [ms]
END_VAR
VAR
    nMs : DINT; // 当日毫秒偏移中间结果 [ms] / intermediate day-millisecond offset [ms]
END_VAR

// 段 1｜返回值与错误状态预置 / segment 1, preset return value and error status
FC_DL_TodToDintMs := DL_TOD_MIN_MS; // 故障缺省返回 0 ms（当日 0 点） [ms] / fault default 0 ms, midnight [ms]
eErr   := 0;     // 预置无错误 / preset no error
bError := FALSE; // 预置无故障（本件无故障级路径） / preset no fault, no fault-level path here
bValid := FALSE; // 预置输出无效，通过域钳位段后置位 / preset invalid, set TRUE after the domain clamp segment

// 段 2｜标准转换链整备 / segment 2, standard conversion chain preparation
nMs := TIME_TO_DINT(TOD_TO_TIME(todIn)); // 标准链：TOD 先转 TIME，再转 DINT 毫秒，绝不自行按时分秒累加 [ms] / standard chain: TOD to TIME then to DINT milliseconds, never accumulate hours/minutes/seconds by hand [ms]

// 段 3｜当日毫秒域钳位（末段） / segment 3, day-millisecond domain clamp (final)
IF nMs < DL_TOD_MIN_MS THEN
    nMs := DL_TOD_MIN_MS; // 越下界钳 0 ms [ms] / clamp upward to 0 ms [ms]
    eErr := 16#0001_01FA; // 信息级：TOD 域外已钳位，正常防御 / info level: out of the TOD domain and clamped, normal defence
ELSIF nMs > DL_TOD_MAX_MS THEN
    nMs := DL_TOD_MAX_MS; // 越上界钳 86399999 ms（24h − 1 ms） [ms] / clamp downward to 86399999 ms, 24h minus 1 ms [ms]
    eErr := 16#0001_01FA; // 同一业务语义复用同一信息码，不另立码 / same business semantics reuses the same info id, no extra code
ELSE
    eErr := 0;            // 域内无错误 / in-domain, no error
END_IF
FC_DL_TodToDintMs := nMs; // 输出钳位后的当日毫秒偏移 [ms] / output the clamped day-millisecond offset [ms]
bError := FALSE;          // 信息级不置故障 / info level never raises fault
bValid := TRUE;           // 域内或钳位后输出均有效可用 / in-domain or clamped output is valid
END_FUNCTION

(* ---- FC_DL_TrapezoidArea.st ---- *)
(*
  ==================================================================
  组件名 Component  : FC_DL_TrapezoidArea
  分类   Category   : DL_MathData
  前缀   Naming     : FC_DL_ ｜ b/n/u/f/t/e/st 类型前缀制（R265）
  复杂度 Complexity  : 低
  版本   Version    : 1.0.0
  功能   Purpose    : 离散序列梯形法累计面积（采样周期入参，纯函数一次算完）。
  来源   Source     : self-std（公开数值积分语义自研包装）
  平台   Platform   : 纯 IEC 61131-3（FOR / 四则 / ABS），三平台通用
  分工声明 Split     : 与 FB_DL_Integrator（连续积分器属主）分工——后者跨拍
                      保持积分状态；本件为无状态纯函数，一次入参一次出面积
                      （R216 双向互引）。
  作者   Author     : 道莅代码库 · PLC 编程专家（R61）
  归属 Ownership     : 本件无 TYPE 声明；引用件类型全部 IEC 标准原生。
  ------------------------------------------------------------------
  边界 Boundary     :
                      一 nCount < 2 无梯形可积：置信息级码、不积累，fArea = 0、
                         bValid = FALSE（信息级不置 bError，R285 口径）；
                      二 采样周期 fDtSec ≤ 0：故障级码，拒绝积分（除法无涉，
                         但零周期等于伪造面积，判故障）；
                      三 NaN 点跳过段计：非有限采样点所在梯形段整段跳过并计数
                         上报 nSkipCnt（信息级，逐点判 x <> x 自反）；
                      四 结果复检兜底同拍置 eErr + bError + bValid 三件套（R258）；
                      五 只读入参数组，不改调用方数据（PercentileLReal 纪律）；
                      六 无状态纯函数：局部量段 1 显式预置（R254）。
  错误码   Codes    :
    16#0001_0633【信息级】采样点数不足（<2），不积累
    16#0001_0634【故障级】采样周期非法（fDtSec ≤ 0），拒绝积分
    16#0001_0635【信息级】存在非有限采样点，已跳过其所在段，个数见 nSkipCnt
    16#0001_0636【故障级】结果非有限（复检兜底）
  验收   Acceptance :
    算法已证（脚本）：未跑 ｜ 编译器已证（三平台）：未跑
    V1 值 0/1/2、fDtSec=1 → 面积 2.0
    V2 nCount=1 → 码 0633、fArea=0、bValid=FALSE
    V3 fDtSec=0 → 码 0634、bError=TRUE
    V4 中间一点 NaN → 码 0635、nSkipCnt=1、有效段照常累加
  修订记录 Revision  :
    2026-11-21  v1.0.0  R61 首版（批 1 · 序号 4）
  ==================================================================
*)
FUNCTION FC_DL_TrapezoidArea : BOOL
VAR_IN_OUT
    afValues : ARRAY[0..1023] OF LREAL; // 采样序列 [工程单位]，前 nCount 个有效 / the sample series, the first nCount entries valid
END_VAR
VAR_INPUT
    nCount  : DINT;  // 采样点数 [个]，合法域 2..1024 / the sample count, legal from two to one thousand twenty four
    fDtSec  : LREAL; // 采样周期 [秒]，必须 > 0 / the sample period in seconds, must be positive
END_VAR
VAR_OUTPUT
    fArea    : LREAL; // 累计面积 [工程单位 × 秒] / the accumulated area
    nSkipCnt : UDINT; // 被跳过的梯形段数 [段] / the skipped trapezoid segment count
    bValid   : BOOL;  // 结果可用标志 [-] / the result usable flag
    eErr     : UDINT; // 错误码，0 = 正常 / the error code, zero is ok
    bError   : BOOL;  // 错误标志，故障级码置位（R45 配对）/ the error flag
END_VAR
VAR
    k        : DINT;  // 段循环索引 [段] / the segment loop index
    nUse     : DINT;  // 钳位后的采样点数 [个] / the clamped sample count
    fV0      : LREAL; // 段左端采样值 [工程单位] / the left sample value of the segment
    fV1      : LREAL; // 段右端采样值 [工程单位] / the right sample value of the segment
    bSkip    : BOOL;  // 本段跳过标记 [-] / the skip flag of this segment
    bClamp   : BOOL;  // 点数钳位标记 [-] / the count clamp flag
END_VAR
VAR CONSTANT
    DL_TRA_NMAX : DINT := 1024; // 采样点容量上界 [个]，与数组容量一致 / the sample capacity aligned with the array
END_VAR

// 段 1｜返回值与错误状态预置安全值（四段式第一段，R45）+ 局部量显式预置（R254）/ segment 1, the preset
FC_DL_TrapezoidArea := FALSE; // 返回值预置假 / preset the return false
fArea := 0.0; // 面积预置零 / preset the area zero
nSkipCnt := 0; // 跳过计数预置零 / preset the skipped count zero
bValid := FALSE; // 有效标志预置假 / preset the validity false
eErr := 16#0000_0000; // 错误码预置正常 / preset the code to ok
bError := FALSE; // 错误标志预置假 / preset the error flag false
nUse := 0; // 采样点数预置零 / preset the count zero
fV0 := 0.0; // 左端值预置零 / preset the left value zero
fV1 := 0.0; // 右端值预置零 / preset the right value zero
bSkip := FALSE; // 跳过标记预置假 / preset the skip flag false
bClamp := FALSE; // 钳位标记预置假 / preset the clamp flag false

// 段 2｜域闸：点数下界早退与上界钳位、周期正域（边界一二）/ segment 2, the count and period gates
IF nCount < 2 THEN // 点数不足：无梯形可积（边界一）/ too few samples, no trapezoid
    eErr := 16#0001_0633; // 信息级：点数不足不积累（信息级不置 bError）/ informational, too few samples
    RETURN; // 早退：fArea 保持零、bValid 保持假 / early return with the area zero
END_IF
IF fDtSec <= 0.0 THEN // 周期非法（边界二）/ an illegal period
    eErr := 16#0001_0634; // 故障级：采样周期非法 / fault grade, the illegal period
    bError := TRUE; // 置错误标志（R45 配对）/ raise the error flag
    bValid := FALSE; // 结果不可用 / the result void
    RETURN; // 早退 / early return
END_IF
nUse := nCount; // 点数域内接管 / take the count
IF nUse > DL_TRA_NMAX THEN // 超容量 / above the capacity
    nUse := DL_TRA_NMAX; // 钳到容量 / clamp to the capacity
    bClamp := TRUE; // 置钳位标记 / raise the clamp flag
END_IF

// 段 3｜梯形法逐段累加（NaN 点整段跳过并计数，边界三）/ segment 3, the segment by segment accumulation with the NaN skip
FOR k := 0 TO nUse - 2 DO // 有界段循环 / the bounded segment loop
    fV0 := afValues[k]; // 左端采样值 / the left sample
    fV1 := afValues[k + 1]; // 右端采样值 / the right sample
    bSkip := (fV0 <> fV0) OR (fV1 <> fV1)
    OR ((fV0 - fV0) <> (fV0 - fV0)) OR ((fV1 - fV1) <> (fV1 - fV1)); // 两端逐点非有限判（NaN 自反 + Inf 差值自减）/ the per point finiteness test
    IF bSkip THEN // 本段含非有限点 / this segment holds a non finite point
        nSkipCnt := nSkipCnt + 1; // 跳过计数推进 / advance the skipped count
    ELSE // 有效段照常累加 / a valid segment accumulates
        fArea := fArea + (fV0 + fV1) * 0.5 * fDtSec; // 梯形面积（除子 2.0 为常量，无除零风险）/ the trapezoid area with a constant divisor
    END_IF
END_FOR

// 段 4｜出口装配：跳过计数与钳位信息级、结果复检兜底（边界四）/ segment 4, the outlet assembly with the recheck
IF nSkipCnt > 0 THEN // 存在被跳过的段 / some segments were skipped
    eErr := 16#0001_0635; // 信息级：非有限点已跳段计数上报 / informational, the skipped segments counted
END_IF
IF (fArea <> fArea) OR ((fArea - fArea) <> (fArea - fArea)) THEN // 结果非有限（结构性不可达兜底）/ the result is not finite, kept as a guard
    fArea := 0.0; // 兜底安全值 / the bottom line safe value
    eErr := 16#0001_0636; // 故障级：结果非有限 / fault grade, the non finite result
    bError := TRUE; // 置错误标志（R45 配对）/ raise the error flag
    bValid := FALSE; // 结果不可用 / the result void
    RETURN; // 早退 / early return
END_IF
bValid := TRUE; // 结果可用 / the result is usable
FC_DL_TrapezoidArea := TRUE; // 返回成功 / return success
END_FUNCTION

(* ---- FC_DL_TrendSlopeCalc.st ---- *)
(*
  FC_DL_TrendSlopeCalc  —  滑窗一阶最小二乘趋势斜率（纯函数）/ Sliding-window least-squares trend slope, pure function
  分类 Category : DL_MathData
  码位 Code     : 16#05_0_04
  段位说明      : 05_0 段仅占 00~03，04/05 为 R38 预留解除后的空穴，本件启用 04 格
  版本 Version  : 1.0.0
  来源 Source   : t2-1-lgf-math — Math 分类「趋势估计」待挖项落地
  溯源 Origin   : clean-room 实现，一阶线性最小二乘为公开经典数学方法，未复制任何源码行
  功能 Function : 1) 对调用方给定的滑窗样本 afY 做一阶最小二乘拟合 y = a + b*x，x = i*fDt；
                  2) 输出斜率 fSlope（趋势速率）、截距 fIntercept、拟合优度 fR2 与有效样本数 nValid；
                  3) 非有限样本（NaN/Inf 判据：x <> x 或幅值越限）自动剔除，不参与拟合；
                  4) 有效样本 < 2、采样间隔 <= 0、SStot 退化为零（常数窗）等边界全部给出确定输出。
  边界 Boundary : ① 纯函数无内部状态，每拍重算；滑窗由调用方持有（FB_DL_SignalStatistics /
                  自管环形窗均可），本件只做一次拟合；
                  ② 与 FB_DL_Differentiator 分工：微分件是瞬时差分、噪声敏感；本件是窗内拟合斜率，
                  供温度升速 / 压降速率 / 泄漏率等趋势判级；
                  ③ 与 FB_DL_*Trend 监视件分工：本件是纯函数估计原子，不做判级、不锁存；
                  ④ 除零守卫：fDt <= 0 直接判无效；SStot 容差判零（浮点禁 = 比较）。
  依赖 Depends  : 无 DL_ 内部依赖，纯 IEC 61131-3
  码表 Error codes（本件格 05_0_04，子码步进 +0x100）:
    16#0005_0104 信息级：非有限样本已剔除（剔后仍 >= 2，拟合照常完成）
    16#0005_0204 故障级：无拟合（有效样本 < 2 或 fDt <= 0 或输入数组非法），返回值 FALSE
    16#0005_0304 信息级：窗内样本为常数（SStot 退化），fR2 置 0，斜率/截距仍有效

  修订历史 Revision :
    2026-11-19  v1.0.0  R39 首版（批次 1 · 序号 2）
*)

FUNCTION FC_DL_TrendSlopeCalc : BOOL    // 返回 TRUE = 拟合有效（斜率/截距/R2 可信）/ TRUE = fit valid
VAR_IN_OUT
    afY : ARRAY[*] OF LREAL;            // 样本窗（时间顺序，最老样本在下标小端）/ Sample window in time order, oldest at low index
END_VAR
VAR_INPUT
    fDt      : LREAL := 1.0;            // 采样间隔 [s]，x = i*fDt，域 > 0 / Sample interval [s], x equals index times fDt
    nCount   : INT := 0;                // 有效样本数声明值 [个]，2..数组维度 / Declared sample count, 2..array size
END_VAR
VAR_OUTPUT
    fSlope     : LREAL;                 // 拟合斜率 b [EU/s]，正值 = 上升趋势 / Fitted slope [EU/s], positive means rising
    fIntercept : LREAL;                 // 拟合截距 a [EU] / Fitted intercept [EU]
    fR2        : LREAL;                 // 拟合优度 R² [无量纲]，0..1，常数窗置 0 / Goodness of fit, 0..1, zero for a constant window
    nValid     : INT;                   // 剔除非有限值后的有效样本数 [个] / Valid sample count after non-finite rejection
    uErrorId   : UDINT;                 // 事件码，0 = 无事件（本件码均为单次调用瞬时，无锁存）/ Event code, transient per call
END_VAR
VAR
    nHi       : INT;                    // 数组上界换算（开放数组） / Resolved array upper bound
    nUse      : INT;                    // 参与拟合的样本数 = MIN(nCount, nHi+1) / Samples actually used
    i         : INT;                    // 遍历索引 / Traversal index
    nGood     : INT;                    // 有限样本计数 [个] / Finite sample counter
    fSumX     : LREAL;                  // Σx 累加器 [s] / Sum of x
    fSumY     : LREAL;                  // Σy 累加器 [EU] / Sum of y
    fSumXY    : LREAL;                  // Σxy 累加器 [EU·s] / Sum of x times y
    fSumX2    : LREAL;                  // Σx² 累加器 [s²] / Sum of x squared
    fDen      : LREAL;                  // 拟合分母 n*Σx² − (Σx)²（前判零）/ Fit denominator, zero-guarded
    fYMean    : LREAL;                  // 有效样本均值 [EU] / Mean of valid samples
    fSStot    : LREAL;                  // 总离差平方和 [EU²] / Total sum of squares
    fSSres    : LREAL;                  // 残差平方和 [EU²] / Residual sum of squares
    fXi       : LREAL;                  // 当前样本横坐标 [s] / Current sample abscissa
    fYi       : LREAL;                  // 当前样本值工作副本 [EU] / Current sample working copy
    fYhat     : LREAL;                  // 当前样本拟合值 [EU] / Fitted value of the current sample
    fDev      : LREAL;                  // 残差工作量 [EU] / Residual working value
END_VAR
VAR CONSTANT
    DL_TSC_N_MIN     : INT   := 2;          // 最少有效样本数 [个] / Minimum valid sample count
    DL_TSC_INF_CAP   : LREAL := 1.0E30;     // 非有限值筛查幅值上限 / Non-finite magnitude screening cap
    DL_TSC_EPS       : LREAL := 1.0E-12;    // 浮点判零容差（分母/SStot 用）/ Float zero tolerance
    DL_TSC_CNT_LIMIT : INT   := 100000;     // nCount 合理上限，防开放数组误传巨大值 / Sane count cap for open arrays
END_VAR

(* —— 段 1｜输出安全预置：任何异常路径下输出必须确定（部分平台残留上次调用值） —— *)
(* Stage 1, safe preset: outputs deterministic on every path *)
FC_DL_TrendSlopeCalc := FALSE;
fSlope     := 0.0;
fIntercept := 0.0;
fR2        := 0.0;
nValid     := 0;
uErrorId   := 16#0005_0204;             // 缺省走「无拟合」故障码，成功路径末尾改写 / Default to no-fit code, rewritten on success

(* —— 段 2｜参数与数组域闸（覆盖参与换算的全部量，R151） —— *)
(* Stage 2, parameter and array gate *)
nHi := UPPER_BOUND(afY, 1) + 1;         // 开放数组元素数 [个] / Element count of the open array
IF nHi < DL_TSC_N_MIN THEN
    RETURN;                             // 数组本身不够两点：无拟合返回 / Array itself too small, return
END_IF
IF fDt <= 0.0 THEN
    RETURN;                             // 采样间隔非法：无拟合返回（防除零口径）
END_IF
nUse := nCount;
IF nUse > nHi THEN
    nUse := nHi;                        // 声明数超过数组维度按维度截断 / Declared count clamped to array size
END_IF
IF nUse > DL_TSC_CNT_LIMIT THEN
    nUse := DL_TSC_CNT_LIMIT;           // 声明数合理上限（防御开放数组误传）/ Sane upper cap
END_IF
IF nUse < DL_TSC_N_MIN THEN
    RETURN;                             // 有效声明样本不足：无拟合返回
END_IF

(* —— 段 3｜单遍累加（剔除非有限样本：x<>x 判 NaN、差值自反判 Inf、幅值兜底） —— *)
(* Stage 3, single pass accumulation with non-finite rejection *)
fSumX  := 0.0;
fSumY  := 0.0;
fSumXY := 0.0;
fSumX2 := 0.0;
nGood  := 0;
FOR i := 0 TO nUse - 1 DO
    fYi := afY[i];                      // 取样本（下标已由 nUse 钳位防越界）/ Fetch sample, index clamped by nUse
    IF (fYi <> fYi) OR (ABS(fYi) > DL_TSC_INF_CAP) OR ((fYi - fYi) <> 0.0) THEN
        uErrorId := 16#0005_0104;       // 信息级：剔除非有限样本（继续累加其余样本）
    ELSE
        fXi   := UDINT_TO_LREAL(UDINT#0 + INT_TO_UDINT(i)) * fDt;   // x = i*fDt（索引先转无符号再乘，防负偏）/ x equals index times fDt
        fSumX  := fSumX  + fXi;
        fSumY  := fSumY  + fYi;
        fSumXY := fSumXY + fXi * fYi;
        fSumX2 := fSumX2 + fXi * fXi;
        nGood  := nGood + 1;
    END_IF
END_FOR
nValid := nGood;
IF nGood < DL_TSC_N_MIN THEN
    RETURN;                             // 有限样本不足：无拟合返回
END_IF

(* —— 段 4｜一阶最小二乘闭式解（分母容差判零，禁 = 号比浮点） —— *)
(* Stage 4, closed-form first-order least squares with zero-guarded denominator *)
fDen := UDINT_TO_LREAL(UDINT#0 + INT_TO_UDINT(nGood)) * fSumX2 - fSumX * fSumX;
IF ABS(fDen) < DL_TSC_EPS THEN
    RETURN;                             // 横坐标退化（窗口时长近零）：无拟合返回
END_IF
fSlope     := (UDINT_TO_LREAL(UDINT#0 + INT_TO_UDINT(nGood)) * fSumXY - fSumX * fSumY) / fDen;   // 斜率（分母已闸）
fIntercept := (fSumY - fSlope * fSumX) / UDINT_TO_LREAL(UDINT#0 + INT_TO_UDINT(nGood));         // 截距（分母 nGood >= 2 恒非零）

(* —— 段 5｜拟合优度 R²（SStot 容差判零；常数窗 R² 置 0 并给信息码） —— *)
(* Stage 5, goodness of fit with degenerate-window guard *)
fYMean := fSumY / UDINT_TO_LREAL(UDINT#0 + INT_TO_UDINT(nGood));
fSStot := 0.0;
fSSres := 0.0;
FOR i := 0 TO nUse - 1 DO
    fYi := afY[i];
    IF (fYi = fYi) AND (ABS(fYi) <= DL_TSC_INF_CAP) AND ((fYi - fYi) = 0.0) THEN   // 仅有效样本参与（与段 3 剔除判据同式）
        fYhat := fIntercept + fSlope * UDINT_TO_LREAL(UDINT#0 + INT_TO_UDINT(i)) * fDt;
        fDev   := fYi - fYhat;
        fSSres := fSSres + fDev * fDev;
        fDev   := fYi - fYMean;
        fSStot := fSStot + fDev * fDev;
    END_IF
END_FOR
IF fSStot < DL_TSC_EPS THEN
    fR2 := 0.0;                         // 常数窗：R² 无定义，置 0，斜率/截距仍有效
    IF uErrorId = 16#0000_0000 THEN
        uErrorId := 16#0005_0304;       // 信息级：常数窗退化（仅在无剔除码时覆盖，剔除码优先保留）
    END_IF
ELSE
    fR2 := 1.0 - fSSres / fSStot;       // R² 换算（分母已闸）
    IF fR2 < 0.0 THEN
        fR2 := 0.0;                     // 数值抖动下限钳位 / Clamp below-zero numerical noise
    END_IF
    IF fR2 > 1.0 THEN
        fR2 := 1.0;                     // 上限钳位 / Upper clamp
    END_IF
END_IF

(* —— 段 6｜成功出口：拟合有效 —— *)
(* Stage 6, success outlet *)
FC_DL_TrendSlopeCalc := TRUE;

END_FUNCTION

(* ---- FC_DL_TriangleSolveSSS.st ---- *)
(*
    FC_DL_TriangleSolveSSS —— SSS 三边解三角形（余弦定理三角度，机构几何 / 三点定位纯函数）
    ------------------------------------------------------------------
    组件名称  : FC_DL_TriangleSolveSSS
    分类      : DL_MathData / Geometry
    前缀      : FC_DL_
    版本      : 1.0.0
    溯源      : 借鉴点 —— 「几何原子归 Math 组」的分类事实（T2-1 Math 行，
                R64 订正遗留的三角方向待挖首件）；余弦定理为公开数学。
                本件无任何 LGF 数据结构 / 命名 / 代码行接触（闭源，只借分类
                事实，最严口径）。
                clean-room 声明 —— 零代码行复制；数学仅用标准运算符与
                ACOS / ABS，域钳位与复验逻辑 100% 自有。
                许可证 —— 本件 MIT。
    平台      : 纯 IEC 61131-3，CODESYS 3.5 / TwinCAT 3 / InoProShop / Machine Expert 通用
    作者      : 道莅代码库 · PLC编程专家（R71 构建轮 · 批 2 · 序号 7）
    ------------------------------------------------------------------
    命名说明  : 泛名 FC_DL_TriangleSolve 在 R71 计划 §2.2 撞名三查中被拒 ——
                与信号发生器 FB_DL_TriangleGenerator（R39 在册）共享
                「Triangle」词根，同根异义高风险命名；故收窄为
                FC_DL_TriangleSolveSSS 并在此声明。本件为 **SSS 专属**
                （三边定三角）：SAS / ASA 等其余解法**不立**（拆件即凑数，
                R62 口径），如有需要由后续轮按独立判据链另行立项。
    功能说明  : 已知三边长（fA / fB / fC，对边对应角 A / B / C），余弦定理
                逐角求解：
                cosA = (b² + c² − a²) / (2·b·c)，A = ACOS(cosA)，B / C 轮换；
                三角和复验 |A + B + C − π| < 1E-6 [rad] 才置返回值 TRUE。
                判据链顺序：三边非有限 / 非正闸 → 三角不等式闸（任意两边
                之和 > 第三边，严格不等；恰等号 = 共线退化 → 拒并出信息码）
                → 余弦定理逐角求解 → 反余弦入参域钳位 [-1, 1]（浮点舍入可致
                比值微越 ±1，直接进 ACOS 得 NaN，R45 口径防域外）→ 三角和
                复验。
                除零面在余弦定理分母 2·b·c：三边非正闸已前置拦截（三边恒正
                则分母恒正），无裸除法暴露；仍做防御性声明（先判后除纪律）。
                浮点判等禁用 =（红线 5）：不等式用严格 > 与容差双口径 ——
                ETOL = 1E-9 [mm] 为绝对容差，仅拦浮点舍入级共线退化
                （工程长度尺度下 1E-9 mm 远小于任何机械可分辨差），域外
                真退化（a + b = c 的实数等号）由严格不等式拒收。
    错误码    : 16#0002_37B0 入参非有限（NaN / Inf / 超幅值）或非正边，角度
                            输出清零 —— 故障级
                16#0002_37B1 三角不等式不成立（含共线退化），拒绝求解，角度
                            输出清零 —— 信息级（几何输入问题，非本件故障）
                16#0002_37B2 三角和复验失败（|Σ−π| >= 1E-6 rad，舍入超差），
                            角度不可信，输出清零 —— 信息级
    码位总账  : 16#0002_37B0 用 ｜ 16#0002_37B1 用 ｜ 16#0002_37B2 用
    状态机    : N/A —— 纯函数无状态，无 CASE 可写，非法状态不可能出现
    边界与披露: 一 无定时器 / 无边沿实例 / 无数组下标，周期安全规则 N/A；
                二 零全局变量、零 VAR_EXTERNAL、零物理地址；
                三 域闸逐项点名（R272）：fA / fB / fC 三入参全部纳入非有限闸
                   （NaN 自反判 + Inf 差值自反判 + 幅值 1E30 上界筛查）与
                   非正闸（<= 0 拒，边长无零边 / 负边语义）；
                四 ACOS 入参钳位 [-1, 1] 必做（浮点舍入可致 > 1），钳位为
                   防御动作不算域外故障，无独立码位（钳后结果仍过三角和
                   复验把守，不静默放行）；
                五 复验失败不置 bError（信息级，R45），返回值 FALSE 即可
                   表达不可信，角度输出一律清零（绝不送未复验值给下游）；
                六 返回值即 bValid 语义（出参契约：三角和复验通过才 TRUE）。
    修订记录  : 2026-11-22 v1.0.0 首次入库（R71 构建轮 · 批 2 · 序号 7）
*)
FUNCTION FC_DL_TriangleSolveSSS : BOOL
VAR_INPUT
    fA : LREAL;                            (* 边长 a（角 A 的对边），[mm]，须 > 0 / the side a, opposite to angle A, must be positive *)
    fB : LREAL;                            (* 边长 b（角 B 的对边），[mm]，须 > 0 / the side b, opposite to angle B, must be positive *)
    fC : LREAL;                            (* 边长 c（角 C 的对边），[mm]，须 > 0 / the side c, opposite to angle C, must be positive *)
END_VAR
VAR_OUTPUT
    fAngA    : LREAL;                      (* 角 A，[rad] / the angle A in radians *)
    fAngB    : LREAL;                      (* 角 B，[rad] / the angle B in radians *)
    fAngC    : LREAL;                      (* 角 C，[rad] / the angle C in radians *)
    nInfoCode: UDINT;                      (* 信息 / 错误码，0 = 正常 / the info or error id, 0 = ok *)
    bError   : BOOL;                       (* 故障标志，仅故障级码置位（R45 配对）/ the fault flag, raised only on fault-level codes *)
END_VAR
VAR CONSTANT
    DL_TSS_FMAX : LREAL := 1.0E30;         (* 非有限筛查幅值上限，[mm] / the finiteness screening cap *)
    DL_TSS_ETOL : LREAL := 1.0E-9;         (* 三角不等式退化容差（绝对口径），[mm] / the degeneracy tolerance of the triangle inequality *)
    DL_TSS_PI   : LREAL := 3.14159265358979; // 圆周率，[rad] / the circle constant pi
    DL_TSS_STOL : LREAL := 1.0E-6;         (* 三角和复验容差，[rad] / the angle sum recheck tolerance *)
END_VAR
VAR
    _fCosA : LREAL;                        (* 角 A 余弦中间量，[无量纲] / the cosine of angle A *)
    _fCosB : LREAL;                        (* 角 B 余弦中间量，[无量纲] / the cosine of angle B *)
    _fCosC : LREAL;                        (* 角 C 余弦中间量，[无量纲] / the cosine of angle C *)
    _fSum  : LREAL;                        (* 三角和中间量，[rad] / the angle sum temporary *)
END_VAR

// 段 1｜返回值与角度预置（统一出口预置，R256）/ segment 1, preset the return and the angles
FC_DL_TriangleSolveSSS := FALSE;           // 故障缺省返回不可信 / the fault default is not trustworthy
fAngA     := 0.0;                          // 角 A 预置零 / preset the angle A to zero
fAngB     := 0.0;                          // 角 B 预置零 / preset the angle B to zero
fAngC     := 0.0;                          // 角 C 预置零 / preset the angle C to zero
nInfoCode := 0;                            // 预置无错 / preset no error
bError    := FALSE;                        // 预置无故障 / preset no fault

// 段 2｜三边非有限闸（NaN 自反判 + Inf 差值自反判 + 幅值上界，R272 逐项点名）/ segment 2, the finiteness gate
IF (fA <> fA) OR ((fA - fA) <> 0.0) OR (ABS(fA) > DL_TSS_FMAX) THEN
    nInfoCode := 16#0002_37B0;             // 故障级：边 a 非有限 / fault level: the side a non finite
    bError := TRUE;                        // R45 配对置故障标志 / paired with the flag
    RETURN;                                // 结构早退（角度保持清零预置）/ structural exit, the angles stay zeroed
END_IF
IF (fB <> fB) OR ((fB - fB) <> 0.0) OR (ABS(fB) > DL_TSS_FMAX) THEN
    nInfoCode := 16#0002_37B0;             // 故障级：边 b 非有限 / fault level: the side b non finite
    bError := TRUE;                        // R45 配对 / paired with the flag
    RETURN;                                // 结构早退 / exit
END_IF
IF (fC <> fC) OR ((fC - fC) <> 0.0) OR (ABS(fC) > DL_TSS_FMAX) THEN
    nInfoCode := 16#0002_37B0;             // 故障级：边 c 非有限 / fault level: the side c non finite
    bError := TRUE;                        // R45 配对 / paired with the flag
    RETURN;                                // 结构早退 / exit
END_IF

// 段 3｜三边非正闸（边长无零边 / 负边语义，兼前置拦余弦定理分母 2·b·c 除零面）/ segment 3, the non positive sides gate
IF (fA <= 0.0) OR (fB <= 0.0) OR (fC <= 0.0) THEN
    nInfoCode := 16#0002_37B0;             // 故障级：非正边 / fault level: a non positive side
    bError := TRUE;                        // R45 配对 / paired with the flag
    RETURN;                                // 结构早退 / exit
END_IF

// 段 4｜三角不等式闸（严格不等 + 容差双口径，恰等号 = 共线退化拒收）/ segment 4, the triangle inequality gate
IF ((fB + fC - fA) <= DL_TSS_ETOL) OR ((fA + fC - fB) <= DL_TSS_ETOL) OR ((fA + fB - fC) <= DL_TSS_ETOL) THEN
    nInfoCode := 16#0002_37B1;             // 信息级：不等式不成立 / info level: the inequality violated
    bError := FALSE;                       // 信息级不置故障（R45）/ info level never raises the flag
    RETURN;                                // 结构早退（角度保持清零）/ exit, the angles stay zeroed
END_IF

// 段 5｜余弦定理逐角求解（分母 2·b·c 已由段 3 前置保证恒正，先判后除纪律已履行）/ segment 5, the cosine theorem per angle
_fCosA := (fB * fB + fC * fC - fA * fA) / (2.0 * fB * fC); // 角 A 余弦 / the cosine of angle A
_fCosB := (fA * fA + fC * fC - fB * fB) / (2.0 * fA * fC); // 角 B 余弦 / the cosine of angle B
_fCosC := (fA * fA + fB * fB - fC * fC) / (2.0 * fA * fB); // 角 C 余弦 / the cosine of angle C

// 段 6｜反余弦入参域钳位 [-1, 1]（浮点舍入防 ACOS 域外 NaN，R45 口径）/ segment 6, the ACOS domain clamp
IF _fCosA > 1.0 THEN                       // 角 A 余弦微越上界 / the cosine slightly over one
    _fCosA := 1.0;                         // 钳到上界 / clamp to one
ELSIF _fCosA < -1.0 THEN                   // 角 A 余弦微越下界 / slightly under minus one
    _fCosA := -1.0;                        // 钳到下界 / clamp to minus one
END_IF
IF _fCosB > 1.0 THEN                       // 角 B 余弦微越上界 / the cosine slightly over one
    _fCosB := 1.0;                         // 钳到上界 / clamp to one
ELSIF _fCosB < -1.0 THEN                   // 角 B 余弦微越下界 / slightly under minus one
    _fCosB := -1.0;                        // 钳到下界 / clamp to minus one
END_IF
IF _fCosC > 1.0 THEN                       // 角 C 余弦微越上界 / the cosine slightly over one
    _fCosC := 1.0;                         // 钳到上界 / clamp to one
ELSIF _fCosC < -1.0 THEN                   // 角 C 余弦微越下界 / slightly under minus one
    _fCosC := -1.0;                        // 钳到下界 / clamp to minus one
END_IF

// 段 7｜反余弦求解（域已钳位，无 NaN 面）/ segment 7, the arccosine solve
fAngA := ACOS(_fCosA);                     // 角 A，[rad] / the angle A
fAngB := ACOS(_fCosB);                     // 角 B，[rad] / the angle B
fAngC := ACOS(_fCosC);                     // 角 C，[rad] / the angle C

// 段 8｜三角和复验（|Σ−π| < 1E-6 rad 才置返回值 TRUE）/ segment 8, the angle sum recheck
_fSum := fAngA + fAngB + fAngC;            // 三角和，[rad] / the angle sum
IF ABS(_fSum - DL_TSS_PI) >= DL_TSS_STOL THEN // 复验失败（舍入超差）/ the recheck failed
    fAngA     := 0.0;                      // 角度不可信，输出清零（绝不送未复验值）/ the angles not trustworthy, zeroed
    fAngB     := 0.0;                      // 清零 / zeroed
    fAngC     := 0.0;                      // 清零 / zeroed
    nInfoCode := 16#0002_37B2;             // 信息级：三角和复验失败 / info level: the recheck failed
    bError    := FALSE;                    // 信息级不置故障（R45）/ info level never raises the flag
    RETURN;                                // 出口（返回值保持 FALSE）/ exit, the return stays FALSE
END_IF

// 段 9｜域内正常出口 / segment 9, the in-domain outlet
FC_DL_TriangleSolveSSS := TRUE;            // 复验通过，角度可信 / the recheck passed, the angles trustworthy
END_FUNCTION
